(* IEC 61131-3 sources: laba_2_/Libraries/Acp10_MC (part 3) *)

FUNCTION_BLOCK MC_BR_OffsetVelocity (*adds a velocity offset to the velocity of the slave axis*)
	VAR_INPUT
		Slave : UDINT; (*axis reference of the slave axis*)
		Enable : BOOL; (*enable the function block*)
		CyclicVelocity : REAL; (*additive velocity*)
		Acceleration : REAL; (*acceleration for reaching the additive velocity*)
		AdvancedParameters : MC_ADV_OFFSETVELOCITY_REF; (*structure for using additional functions*)
	END_VAR
	VAR_OUTPUT
		Active : BOOL; (*a velocity offset can be executed*)
		Busy : BOOL; (*function block is not finished*)
		Error : BOOL; (*error occurred in FB*)
		ErrorID : UINT; (*error number*)
		VelocityAttained : BOOL; (*additive velocity offset reached*)
		ActualShiftValue : REAL; (*current value of velocity offset on the drive*)
	END_VAR
	VAR
		C_Slave : UDINT; (*internal variable*)
		IS : MC_0127_IS_TYP; (*internal variable*)
	END_VAR
END_FUNCTION_BLOCK

FUNCTION_BLOCK MC_BR_OffsetZone (*adds an offset to the position of the slave axis*)
	VAR_INPUT
		Slave : UDINT; (*axis reference of the slave axis*)
		Enable : BOOL; (*enable the function block*)
		InitData : BOOL; (*initialize the input data*)
		Shift : REAL; (*offset shift value*)
		Velocity : REAL; (*velocity for reaching the offset shift*)
		Acceleration : REAL; (*acceleration for reaching the offset shift*)
		ZoneStartPosition : REAL; (*start position of the offset shift zone*)
		ZoneEndPosition : REAL; (*end position of the offset shift zone*)
		AdvancedParameters : MC_ADV_OFFSETZONE_REF; (*structure for using additional functions*)
	END_VAR
	VAR_OUTPUT
		Active : BOOL; (*a offset shift can be executed*)
		Busy : BOOL; (*function block is not finished*)
		Error : BOOL; (*error occurred in FB*)
		ErrorID : UINT; (*error number*)
		ShiftAttained : BOOL; (*offset shift executed*)
		DataInitialized : BOOL; (*input data initialized*)
		ActualShiftValue : REAL; (*current value of shift on the drive*)
	END_VAR
	VAR
		C_Slave : UDINT; (*internal variable*)
		IS : MC_0128_IS_TYP; (*internal variable*)
	END_VAR
END_FUNCTION_BLOCK

FUNCTION_BLOCK MC_BR_GetParIDInfo (*determines data type and data length of a ParID*)
	VAR_INPUT
		Execute : BOOL; (*determine ParID information at rising edge*)
		ParID : UINT; (*ParID of which the information should be determined*)
	END_VAR
	VAR_OUTPUT
		Done : BOOL; (*command executed*)
		Busy : BOOL; (*function block is not finished*)
		Error : BOOL; (*error occurred in FB*)
		ErrorID : UINT; (*error number*)
		ParIDInfo : MC_PARID_INFO_REF; (*information about ParID*)
	END_VAR
	VAR
		IS : MC_0106_IS_TYP; (*intern variable*)
	END_VAR
END_FUNCTION_BLOCK

FUNCTION_BLOCK MC_BR_ParTrace (*controls the parameter trace*)
	VAR_INPUT
		Execute : BOOL; (*execute command at rising edge*)
		Command : UINT; (*select the command for the trace*)
		Configuration : MC_PARTRACECONFIG_REF; (*FB configuration*)
	END_VAR
	VAR_OUTPUT
		Done : BOOL; (*command executed*)
		Busy : BOOL; (*function block is not finished*)
		Error : BOOL; (*error occurred in FB*)
		ErrorID : UINT; (*error number*)
		ErrorRecord : MC_ERRORRECORD_REF; (*error messages that can occur after executing the command*)
	END_VAR
	VAR
		IS : MC_0080_IS_TYP; (*intern variable*)
	END_VAR
END_FUNCTION_BLOCK

FUNCTION_BLOCK MC_BR_ParTraceConfig (*load and save axis trace configuration*)
	VAR_INPUT
		Execute : BOOL; (*execute command at rising edge*)
		Command : UINT; (*select the command for the trace*)
		AdrTraceConfig : UDINT; (*adress of axis trace configuration*)
		DataObject : MC_DATOBJ_REF; (*data object parameters*)
	END_VAR
	VAR_OUTPUT
		Done : BOOL; (*command executed*)
		Busy : BOOL; (*function block is not finished*)
		Error : BOOL; (*error occurred in FB*)
		ErrorID : UINT; (*error number*)
		ErrorRecord : MC_ERRORRECORD_REF; (*error messages that can occur after executing the command*)
	END_VAR
	VAR
		IS : MC_0102_IS_TYP; (*intern variable*)
	END_VAR
END_FUNCTION_BLOCK

FUNCTION_BLOCK MC_BR_Phasing (*causes a phase shift in the master position of the slave axis*)
	VAR_INPUT
		Slave : UDINT; (*axis reference of the slave axis*)
		Enable : BOOL; (*enable the function block*)
		InitData : BOOL; (*initialize the input data*)
		PerformVelocityControl : BOOL; (*enable the phase shift*)
		Shift : REAL; (*phase shift value*)
		Velocity : REAL; (*velocity for reaching the phase shift*)
		Acceleration : REAL; (*acceleration for reaching the phase shift*)
		ApplicationDistance : REAL; (*distance within which the phase shift occurs*)
		ApplicationMode : UINT; (*basis for movement profile*)
		ShiftMode : UINT; (*definition of how the value on the "Shift" input should be used*)
		AdvancedParameters : MC_ADVANCEDSHIFTPAR_REF; (*structure for using additional functions*)
	END_VAR
	VAR_OUTPUT
		Active : BOOL; (*a phase shift can be executed*)
		Busy : BOOL; (*function block is not finished*)
		Error : BOOL; (*error occurred in FB*)
		ErrorID : UINT; (*error number*)
		ShiftAttained : BOOL; (*phase shift executed*)
		DataInitialized : BOOL; (*input data initialized*)
		ActualShiftValue : REAL; (*current value of shift on the drive*)
	END_VAR
	VAR
		C_Slave : UDINT; (*internal variable*)
		C_InitData : BOOL; (*internal variable*)
		C_PerformVelocityControl : BOOL; (*internal variable*)
		C_Shift : DINT; (*internal variable*)
		C_Velocity : REAL; (*internal variable*)
		C_Acceleration : REAL; (*internal variable*)
		C_ApplicationDistance : DINT; (*internal variable*)
		C_ApplicationMode : UINT; (*internal variable*)
		C_SelectedMaster : UINT; (*internal variable*)
		C_ShiftMode : UINT; (*internal variable*)
		C_AdvancedParameters : MC_ADVANCEDSHIFTPAR_REF; (*internal variable*)
		C_Active : BOOL; (*internal variable*)
		C_Busy : BOOL; (*internal variable*)
		C_Error : BOOL; (*internal variable*)
		C_ErrorID : UINT; (*internal variable*)
		CC_ErrorID : UINT; (*internal variable*)
		C_ShiftAttained : BOOL; (*internal variable*)
		C_DataInitialized : BOOL; (*internal variable*)
		C_AxisState : UINT; (*internal variable*)
		NextState : USINT; (*internal variable*)
		state : USINT; (*internal variable*)
		LockID : USINT; (*internal variable*)
		LockIDPar : USINT; (*internal variable*)
		Factor : UDINT; (*internal variable*)
		RtN : REAL; (*internal variable*)
		VarIndex : UINT; (*internal variable*)
		MpgenIndex : UINT; (*internal variable*)
		C_MpgenStatus : USINT; (*internal variable*)
		MpgenStatusOffset : UINT; (*internal variable*)
		MpgenStatusRecIndex : USINT; (*internal variable*)
		Reserve : USINT; (*internal variable*)
		MpgenValueOffset : UINT; (*internal variable*)
		MpgenValueRecIndex : USINT; (*internal variable*)
		FbID : USINT; (*internal variable*)
		InitDataActive : BOOL; (*internal variable*)
	END_VAR
END_FUNCTION_BLOCK

FUNCTION_BLOCK MC_BR_MechPosDeviationComp (*handles mechanics position deviation compensation*)
	VAR_INPUT
		Axis : UDINT; (*axis reference*)
		Enable : BOOL; (*as long as Enable is TRUE the FB is active*)
		Parameters : MC_MPDC_PARAM_REF; (*parameters for mechanics position deviation compensation*)
		AdvancedParameters : MC_ADV_MPDC_REF; (*advanced parameters for mechanics deviation position compensation*)
	END_VAR
	VAR_OUTPUT
		Active : BOOL; (*if set, the mechanics deviation position compensation is active*)
		Busy : BOOL; (*function block is not finished*)
		Error : BOOL; (*error occurred in FB*)
		ErrorID : UINT; (*error number*)
		AdvancedInfo : MC_ADV_INFO_MPDC_REF; (*structure with additional information*)
	END_VAR
	VAR
		C_Axis : UDINT; (*internal variable*)
		IS : MC_0147_IS_TYP; (*internal structure*)
	END_VAR
END_FUNCTION_BLOCK

FUNCTION_BLOCK MC_BR_PowerMeter (*executes the evaluation of the powerdata of a PSM*)
	VAR_INPUT
		Axis : UDINT; (*axis reference*)
		Enable : BOOL; (*as long as Enable is TRUE the power evaluation is active*)
		Mode : USINT; (*choose the mode for the power evaluation*)
		IntervalTime : UINT; (*duration of the interval*)
		RestartInterval : BOOL; (*a new interval is startet at rising edge of this input*)
		EventInput : MC_BR_EVINPUT_REF; (*if this is used, the Trigger input will not be considered*)
	END_VAR
	VAR_OUTPUT
		Valid : BOOL; (*if set, the data on Output PowerData are valid*)
		Busy : BOOL; (*function block is not finished*)
		Error : BOOL; (*error occurred in FB*)
		ErrorID : UINT; (*error number*)
		PowerData : MC_POWERDATA_REF; (*structure for the power data*)
		MissedIntervals : UINT; (*count of missed intervalls*)
	END_VAR
	VAR
		C_Axis : UDINT; (*internal variable*)
		IS : MC_0089_IS_TYP; (*internal structure*)
	END_VAR
END_FUNCTION_BLOCK

FUNCTION_BLOCK MC_BR_ReadAutPosition (*reads the cam profile automat position*)
	VAR_INPUT
		Axis : UDINT; (*axis reference*)
		Execute : BOOL; (*automat position is read at rising edge*)
	END_VAR
	VAR_OUTPUT
		Done : BOOL; (*reading automat position is finished*)
		Busy : BOOL; (*function block is not finished*)
		Error : BOOL; (*error occurred in FB*)
		ErrorID : UINT; (*error number*)
		AutPosition : REAL; (*automat position*)
	END_VAR
	VAR
		C_Axis : UDINT; (*internal variable*)
		C_Execute : BOOL; (*internal variable*)
		C_Done : BOOL; (*internal variable*)
		C_Error : BOOL; (*internal variable*)
		C_ErrorID : UINT; (*internal variable*)
		LockIDPar : USINT; (*internal variable*)
		Reserve1 : USINT; (*internal variable*)
		C_AutPosition : DINT; (*internal variable*)
		C_DataAddress : UDINT; (*internal variable*)
		state : USINT; (*internal variable*)
	END_VAR
END_FUNCTION_BLOCK

FUNCTION_BLOCK MC_BR_ReadAxisError (*reads and acknowledges an axis error record and reads the error text*)
	VAR_INPUT
		Axis : UDINT; (*axis reference*)
		Enable : BOOL; (*read error record/text*)
		Acknowledge : BOOL; (*acknowledge current axis error*)
		Mode : UINT; (*operating mode of FB*)
		Configuration : MC_ERRORTEXTCONFIG_REF; (*FB configuration*)
	END_VAR
	VAR_OUTPUT
		Valid : BOOL; (*if set, the data of the other outputs is valid*)
		Busy : BOOL; (*function block is not finished*)
		Error : BOOL; (*error occurred in FB*)
		ErrorID : UINT; (*error number*)
		ErrorRecordAvailable : BOOL; (*a new error record is available*)
		ErrorRecord : MC_ERRORRECORD_REF; (*detailed axis error information*)
		FunctionBlockErrorCount : UINT; (*number of not acknowledged function block errors*)
		AxisErrorCount : UINT; (*number of not acknowledged axis errors*)
		AxisWarningCount : UINT; (*number of not acknowledged axis warnings*)
	END_VAR
	VAR
		C_Axis : UDINT; (*internal variable*)
		IS : MC_0105_IS_TYP; (*internal variable*)
	END_VAR
END_FUNCTION_BLOCK

FUNCTION_BLOCK MC_BR_ReadCyclicPosition (*read the position of an axis cyclically*)
	VAR_INPUT
		Axis : UDINT; (*axis reference*)
		Enable : BOOL; (*as long as Enable is TRUE the cyclic position is read from the axis*)
		ParID : UINT; (*ParID that is read cyclically, 0... set position*)
	END_VAR
	VAR_OUTPUT
		Valid : BOOL; (*position is beeing read from the axis*)
		Busy : BOOL; (*function block is not finished*)
		Error : BOOL; (*error occurred in FB*)
		ErrorID : UINT; (*error number*)
		CyclicPosition : MC_CYCLIC_POSITION; (*cyclic position that is read from the axis*)
	END_VAR
	VAR
		C_Axis : UDINT; (*internal variable*)
		IS : MC_0082_IS_TYP; (*internal variable*)
	END_VAR
END_FUNCTION_BLOCK

FUNCTION_BLOCK MC_BR_ReadDriveStatus (*checks the status of a drive*)
	VAR_INPUT
		Axis : UDINT; (*axis reference*)
		Enable : BOOL; (*when set the status is read*)
		AdrDriveStatus : UDINT; (*address of the structur where the status is written on*)
	END_VAR
	VAR_OUTPUT
		Valid : BOOL; (*output of FB is valid*)
		Busy : BOOL; (*function block is not finished*)
		Error : BOOL; (*error occurred in FB*)
		ErrorID : UINT; (*error number*)
	END_VAR
	VAR
		C_Axis : UDINT; (*internal variable*)
		state : USINT; (*internal variable*)
		C_Error : BOOL; (*internal variable*)
		C_ErrorID : UINT; (*internal variable*)
		C_AdrDriveStatus : UDINT; (*internal variable*)
	END_VAR
END_FUNCTION_BLOCK

FUNCTION_BLOCK MC_BR_ReadNetTraceStatus (*determines the current status of the network command trace*)
	VAR_INPUT
		Enable : BOOL; (*the status of the network command trace is read as long as the input is enabled*)
		Configuration : MC_NETTRACECONFIG_REF; (*FB configuration. Only the element "NetTrace" is evaluated*)
	END_VAR
	VAR_OUTPUT
		Valid : BOOL; (*the status information is valid*)
		Busy : BOOL; (*function block is not finished*)
		Error : BOOL; (*error occurred in FB*)
		ErrorID : UINT; (*error number*)
		TraceState : UINT; (*status of the NWCT*)
	END_VAR
	VAR
		C_ErrorID : UINT; (*internal variable*)
		C_Error : BOOL; (*internal variable*)
		state : USINT; (*internal variable*)
	END_VAR
END_FUNCTION_BLOCK

FUNCTION_BLOCK MC_BR_ReadParID (*reads a ParID from the specified axis*)
	VAR_INPUT
		Axis : UDINT; (*axis reference*)
		Execute : BOOL; (*read data at rising edge*)
		ParID : UINT; (*number of the parameter ID to read*)
		DataAddress : UDINT; (*address of the user variable*)
		DataType : UINT; (*data type of the user variable*)
	END_VAR
	VAR_OUTPUT
		Done : BOOL; (*value of ParID has been copied to the user variable*)
		Busy : BOOL; (*function block is not finished*)
		Error : BOOL; (*error occurred in function block*)
		ErrorID : UINT; (*error number*)
	END_VAR
	VAR
		C_Axis : UDINT; (*internal variable*)
		C_Execute : BOOL; (*internal variable*)
		C_ParID : UINT; (*internal variable*)
		LockIDPar : USINT; (*internal variable*)
		Reserve1 : USINT; (*internal variable*)
		C_DataAddress : UDINT; (*internal variable*)
		Reserve2 : UDINT; (*internal variable*)
		C_DataType : UINT; (*internal variable*)
		C_Done : BOOL; (*internal variable*)
		C_Error : BOOL; (*internal variable*)
		C_ErrorID : UINT; (*internal variable*)
		state : USINT; (*internal variable*)
	END_VAR
END_FUNCTION_BLOCK

FUNCTION_BLOCK MC_BR_ReadParIDText (*reads a ParID from the specified axis in text format*)
	VAR_INPUT
		Axis : UDINT; (*axis reference*)
		Execute : BOOL; (*read data at rising edge*)
		ParID : UINT; (*number of the parameter ID to read*)
	END_VAR
	VAR_OUTPUT
		Done : BOOL; (*value of ParID has been read*)
		Busy : BOOL; (*function block is not finished*)
		Error : BOOL; (*error occurred in function block*)
		ErrorID : UINT; (*error number*)
		DataText : STRING[33]; (*value of ParID in text format *)
	END_VAR
	VAR
		C_Axis : UDINT; (*internal variable*)
		C_Execute : BOOL; (*internal variable*)
		C_ParID : UINT; (*internal variable*)
		LockIDPar : USINT; (*internal variable*)
		C_Done : BOOL; (*internal variable*)
		C_Error : BOOL; (*internal variable*)
		C_ErrorID : UINT; (*internal variable*)
		state : USINT; (*internal variable*)
	END_VAR
END_FUNCTION_BLOCK

FUNCTION_BLOCK MC_BR_ReadParList (*read a parameter list*)
	VAR_INPUT
		Axis : UDINT; (*axis reference*)
		Execute : BOOL; (*read parameter list at rising edge*)
		DataAddress : UDINT; (*address of the parameter list*)
	END_VAR
	VAR_OUTPUT
		Done : BOOL; (*transfer completed*)
		Busy : BOOL; (*function block is not finished*)
		Error : BOOL; (*error occurred in FB*)
		ErrorID : UINT; (*error number*)
	END_VAR
	VAR
		LockIDPar : USINT; (*internal variable*)
		C_Error : BOOL; (*internal variable*)
		C_ErrorID : UINT; (*internal variable*)
		C_Axis : UDINT; (*internal variable*)
		C_DataAddress : UDINT; (*internal variable*)
		C_Done : BOOL; (*internal variable*)
		state : USINT; (*internal variable*)
	END_VAR
END_FUNCTION_BLOCK

FUNCTION_BLOCK MC_BR_ReadParTraceStatus (*determines the current status of the axis trace*)
	VAR_INPUT
		Enable : BOOL; (*the status of the axis trace is read as long as the input is enabled*)
		Configuration : MC_PARTRACECONFIG_REF; (*FB configuration. Only the element "ParTrace" is evaluated*)
	END_VAR
	VAR_OUTPUT
		Valid : BOOL; (*the status information is valid*)
		Busy : BOOL; (*function block is not finished*)
		Error : BOOL; (*error occurred in FB*)
		ErrorID : UINT; (*error number*)
		TraceState : UINT; (*status of the trace*)
	END_VAR
	VAR
		C_ErrorID : UINT; (*internal variable*)
		C_Error : BOOL; (*internal variable*)
		state : USINT; (*internal variable*)
	END_VAR
END_FUNCTION_BLOCK

FUNCTION_BLOCK MC_BR_ReceiveParIDOnPLC (*initializes receiving of a ParID on the PLC*)
	VAR_INPUT
		Axis : UDINT; (*axis reference*)
		Enable : BOOL; (*as long as Enable is TRUE the ParID is read from the axis*)
		ParID : UINT; (*ParID that is read cyclically*)
		SendChannel : USINT; (*send channel on which the ParID is sent*)
		Mode : USINT; (*convertion of ParID-value into PLCopen-units can be activated*)
	END_VAR
	VAR_OUTPUT
		Valid : BOOL; (*ParID is beeing read from the axis*)
		Busy : BOOL; (*function block is not finished*)
		Error : BOOL; (*error occurred in FB*)
		ErrorID : UINT; (*error number*)
		CyclicValue : MC_CYCLIC_VALUE_REF; (*cyclic ParID value that is read from the axis*)
	END_VAR
	VAR
		C_Axis : UDINT; (*internal variable*)
		IS : MC_0113_IS_TYP; (*internal variable*)
	END_VAR
END_FUNCTION_BLOCK

FUNCTION_BLOCK MC_BR_ResetAutPar (*initializes the general parameters of the cam automat*)
	VAR_INPUT
		Axis : UDINT; (*axis reference*)
		Execute : BOOL; (*set parameter to default values at rising edge*)
		GlobalParams : USINT; (*selection of the global parameter*)
		StateIndex : USINT; (*selection of the automat state*)
	END_VAR
	VAR_OUTPUT
		Done : BOOL; (*automat parameters set to default values*)
		Busy : BOOL; (*function block not finished*)
		Error : BOOL; (*error occurred in FB*)
		ErrorID : UINT; (*error number*)
	END_VAR
	VAR
		C_Axis : UDINT; (*internal variable*)
		IS : MC_0136_IS_TYP; (*internal variable*)
	END_VAR
END_FUNCTION_BLOCK

FUNCTION_BLOCK MC_BR_SaveAxisPar (*writes the axis parameters in the axis data structure*)
	VAR_INPUT
		Axis : UDINT; (*axis reference*)
		Execute : BOOL; (*write axis parameter from the axis structure to a init parameter module at rising edge*)
		DataObjectName : STRING[12]; (*name of the init parameter module*)
	END_VAR
	VAR_OUTPUT
		Done : BOOL; (*saving the data is finished*)
		Busy : BOOL; (*function block is not finished*)
		Error : BOOL; (*error occurred in FB*)
		ErrorID : UINT; (*error number*)
		DataObjectIdent : UDINT; (*init parameter module data object ID for the function blocks in the DataObj library*)
	END_VAR
	VAR
		C_Axis : UDINT;
		C_DataObjectName : STRING[12]; (*internal variable*)
		state : USINT; (*internal variable*)
		LockIDPar : USINT; (*internal variable*)
		C_ErrorID : UINT; (*internal variable*)
		C_Error : BOOL; (*internal variable*)
		pInit : REFERENCE TO USINT; (*internal variable*)
		pError : REFERENCE TO USINT; (*internal variable*)
	END_VAR
END_FUNCTION_BLOCK

FUNCTION_BLOCK MC_BR_SaveCamProfileObj (*saves the data of a cam profile into a data module*)
	VAR_INPUT
		Execute : BOOL; (*save the cam profile at rising edge*)
		DataObjectName : STRING[12]; (*name for the data module in which the cam profile is saved*)
		DataAddress : UDINT; (*address of the cam profile data*)
		DataObjectVersion : UINT; (*version for the data module*)
	END_VAR
	VAR_OUTPUT
		Done : BOOL; (*data module was saved*)
		Busy : BOOL; (*function block is not finished*)
		Error : BOOL; (*error occurred in FB*)
		ErrorID : UINT; (*error number*)
		ErrorRecord : MC_ERRORRECORD_REF; (*error messages that can occur after executing the command*)
		DataObjectIdent : UDINT; (*ident of the data module*)
	END_VAR
	VAR
		IS : MC_0116_IS_TYP; (*internal variable*)
	END_VAR
END_FUNCTION_BLOCK

FUNCTION_BLOCK MC_BR_SetHardwareInputs (*forces the hardware inputs*)
	VAR_INPUT
		Axis : UDINT; (*axis reference*)
		Enable : BOOL; (*set the status of the hardware inputs as long as the input is enabled*)
		HomeSwitch : BOOL; (*if TRUE the reference hardware input is activated*)
		PosHWSwitch : BOOL; (*if TRUE the positive limit switch input is activated*)
		NegHWSwitch : BOOL; (*if TRUE the negative limit switch input is activated*)
		Trigger1 : BOOL; (*if TRUE the trigger1 input is activated*)
		Trigger2 : BOOL; (*if TRUE the trigger2 input is activated*)
	END_VAR
	VAR_OUTPUT
		Active : BOOL; (*function block is active and waits for changes on the inputs*)
		Busy : BOOL; (*function block is not finished*)
		Error : BOOL; (*error occurred in FB*)
		ErrorID : UINT; (*error number*)
		InputsSet : BOOL; (*the actual input status was transferred*)
	END_VAR
	VAR
		C_Axis : UDINT; (*internal variable*)
		IS : MC_0108_IS_TYP; (*internal variable*)
	END_VAR
END_FUNCTION_BLOCK

FUNCTION_BLOCK MC_BR_SetupController (*starts a controller setup and saves the parameters*)
	VAR_INPUT
		Axis : UDINT; (*axis reference*)
		Execute : BOOL; (*starts the command action at rising edge*)
		Command : UINT; (*choose the command for the setup*)
		Configuration : MC_SETUP_CONTROLLER_CFG_REF; (*FB-Configuration*)
	END_VAR
	VAR_OUTPUT
		Done : BOOL; (*command successfully completed*)
		Busy : BOOL; (*function block is not finished*)
		CommandAborted : BOOL; (*function block is aborted by another command*)
		Error : BOOL; (*error occurred in FB*)
		ErrorID : UINT; (*error number*)
		SetupOutput : MC_SETUP_OUTPUT_REF; (*structure for output values*)
	END_VAR
	VAR
		C_Axis : UDINT; (*internal variable*)
		IS : MC_0090_IS_TYP; (*internal variable*)
	END_VAR
END_FUNCTION_BLOCK

FUNCTION_BLOCK MC_BR_SetupFromParTabObj (*starts a setup with parameter from an ACOPOS parameter table*)
	VAR_INPUT
		Axis : UDINT; (*axis reference*)
		Execute : BOOL; (*starts the commanded action at rising edge*)
		Command : UINT; (*choose the command for the setup*)
		DataObjectName : STRING[12]; (*name of the ACOPOS parameter table*)
	END_VAR
	VAR_OUTPUT
		Done : BOOL; (*command succesfully completed*)
		Busy : BOOL; (*function block is not finished*)
		CommandAborted : BOOL; (*function block is aborted by another command*)
		Error : BOOL; (*error occurred in FB*)
		ErrorID : UINT; (*error number*)
		SetupOutput : MC_SETUP_OUTPUT_REF; (*structure for output values*)
	END_VAR
	VAR
		C_Axis : UDINT; (*internal variable*)
		IS : MC_0145_IS_TYP; (*internal variable*)
	END_VAR
END_FUNCTION_BLOCK

FUNCTION_BLOCK MC_BR_SetupInductionMotor (*starts the motorsetup for an induction motor and saves the parameters*)
	VAR_INPUT
		Axis : UDINT; (*axis reference*)
		Execute : BOOL; (*starts the commanded action at rising edge*)
		Command : UINT; (*choose the command for the setup*)
		Configuration : MC_SETUP_IND_MOTOR_CFG_REF; (*FB-Configuration*)
	END_VAR
	VAR_OUTPUT
		Done : BOOL; (*command succesfully completed*)
		Busy : BOOL; (*function block is not finished*)
		CommandAborted : BOOL; (*function block is aborted by another command*)
		Error : BOOL; (*error occurred in FB*)
		ErrorID : UINT; (*error number*)
		SetupOutput : MC_SETUP_OUTPUT_REF; (*structure for output values*)
	END_VAR
	VAR
		C_Axis : UDINT; (*internal variable*)
		IS : MC_0088_IS_TYP; (*internal variable*)
	END_VAR
END_FUNCTION_BLOCK

FUNCTION_BLOCK MC_BR_SetupIsqRipple (*starts the setup for isq ripple compensation  and saves the parameters*)
	VAR_INPUT
		Axis : UDINT; (*axis reference*)
		Execute : BOOL; (*starts the commanded action at rising edge*)
		Command : UINT; (*choose the command for the setup*)
		Configuration : MC_SETUP_ISQ_RIPPLE_CFG_REF; (*FB-Configuration*)
	END_VAR
	VAR_OUTPUT
		Done : BOOL; (*command successfully completed*)
		Busy : BOOL; (*function block is not finished*)
		CommandAborted : BOOL; (*function block is aborted by another command*)
		Error : BOOL; (*error occurred in FB*)
		ErrorID : UINT; (*error number*)
		SetupOutput : MC_SETUP_OUTPUT_REF; (*structure for the output values*)
	END_VAR
	VAR
		C_Axis : UDINT; (*internal variable*)
		IS : MC_0101_IS_TYP; (*internal variable*)
	END_VAR
END_FUNCTION_BLOCK

FUNCTION_BLOCK MC_BR_SetupMotorPhasing (*starts a phasing setup and saves the parameters*)
	VAR_INPUT
		Axis : UDINT; (*axis reference*)
		Execute : BOOL; (*starts the commanded action at rising edge*)
		Command : UINT; (*choose the command for the setup*)
		Configuration : MC_SETUP_MOTOR_PHA_CFG_REF; (*FB-Configuration*)
	END_VAR
	VAR_OUTPUT
		Done : BOOL; (*command successfully completed*)
		Busy : BOOL; (*function block is not finished*)
		CommandAborted : BOOL; (*function block is aborted by another command*)
		Error : BOOL; (*error occurred in FB*)
		ErrorID : UINT; (*error number *)
		SetupOutput : MC_SETUP_OUTPUT_REF; (*structure for output values*)
		SetupResult : MC_SETUP_PHASING_RESULT_REF; (*structure for results of the setup*)
	END_VAR
	VAR
		C_Axis : UDINT; (*internal variable*)
		IS : MC_0097_IS_TYP; (*internal variable*)
	END_VAR
END_FUNCTION_BLOCK

FUNCTION_BLOCK MC_BR_SetupSynchronMotor (*starts the motorsetup for a synchron motor and saves the parameters*)
	VAR_INPUT
		Axis : UDINT; (*axis reference*)
		Execute : BOOL; (*starts the commanded action at rising edge*)
		Command : UINT; (*choose the command for the setup*)
		Configuration : MC_SETUP_SYNC_MOTOR_CFG_REF; (*FB-Configuration*)
	END_VAR
	VAR_OUTPUT
		Done : BOOL; (*command successfully completed*)
		Busy : BOOL; (*function block is not finished*)
		CommandAborted : BOOL; (*function block is aborted by another command*)
		Error : BOOL; (*error occurred in FB*)
		ErrorID : UINT; (*error number*)
		SetupOutput : MC_SETUP_OUTPUT_REF; (*structure for output values*)
	END_VAR
	VAR
		C_Axis : UDINT; (*internal variable*)
		IS : MC_0129_IS_TYP; (*internal variable*)
	END_VAR
END_FUNCTION_BLOCK

FUNCTION_BLOCK MC_BR_Simulation (*turns on or off simulation mode for a drive*)
	VAR_INPUT
		Axis : UDINT; (*axis reference*)
		Execute : BOOL; (*switch simulation mode on or off at rising edge*)
		SimulationCommand : UINT; (*choose if switch on or off simulation mode*)
	END_VAR
	VAR_OUTPUT
		Done : BOOL; (*simulation mode is on or off*)
		Busy : BOOL; (*function block is not finished*)
		Error : BOOL; (*error occurred in FB*)
		ErrorID : UINT; (*error number*)
	END_VAR
	VAR
		C_Axis : UDINT; (*internal variable*)
		IS : MC_0071_IS_TYP; (*internal variable*)
	END_VAR
END_FUNCTION_BLOCK

FUNCTION_BLOCK MC_BR_TouchProbe (*saves the values of ParIDs when a specified event occurs*)
	VAR_INPUT
		Axis : UDINT; (*axis reference*)
		TriggerInput : MC_BR_TRIGGER_REF; (*input that is used as event source*)
		Enable : BOOL; (*as long as enable is TRUE, a value is saved every time a trigger event occurs*)
		Period : REAL; (*interval between two expected trigger positions*)
		PeriodChange : REAL; (*if no valid event occurs within an interval, the window is shifted by the value of Period*)
		ExpectedValue : REAL; (*expected position of the trigger event within the Period*)
		WindowNegative : REAL; (*range before the expected position in which the trigger signal may occur*)
		WindowPositive : REAL; (*range after the expected position in which the trigger signal may occur*)
		Mode : UINT; (*the way the FB works can be determined with this input*)
	END_VAR
	VAR_OUTPUT
		Active : BOOL; (*waits for a trigger event*)
		Busy : BOOL; (*function block is not finished*)
		Error : BOOL; (*error occured in FB*)
		ErrorID : UINT; (*error number*)
		RecordedPeriodicValue : REAL; (*result value within the configured period*)
		RecordedValue : DINT; (*result value*)
		DeltaExpectedValue : REAL; (*deviation: expected position - result value*)
		ProbeCounter : UDINT; (*number of valid trigger events since "Enable" was set to TRUE*)
		MissedTriggers : UDINT; (*number of invalid or missing trigger events since "Enable" was set to TRUE*)
	END_VAR
	VAR
		C_Axis : UDINT; (*internal variable*)
		C_TriggerInput : MC_BR_TRIGGER_REF; (*internal variable*)
		C_Period : DINT; (*internal variable*)
		C_PeriodChange : DINT; (*internal variable*)
		C_ExpectedValue : DINT; (*internal variable*)
		C_WindowNegative : DINT; (*internal variable*)
		C_WindowPositive : DINT; (*internal variable*)
		C_Mode : UINT; (*internal variable*)
		C_Active : BOOL; (*internal variable*)
		C_Busy : BOOL; (*internal variable*)
		C_Error : BOOL; (*internal variable*)
		C_ErrorID : UINT; (*internal variable*)
		C_RecordedPeriodicValue : REAL; (*internal variable*)
		C_RecordedValue : DINT; (*internal variable*)
		C_DeltaExpectedValue : REAL; (*internal variable*)
		C_ProbeCounter : UDINT; (*internal variable*)
		C_MissedTriggers : UDINT; (*internal variable*)
		PeriodOffset : DINT; (*internal variable*)
		LatchValue : DINT; (*internal variable*)
		LatchDeltaIv : DINT; (*internal variable*)
		NewValue : BOOL; (*internal variable*)
		state : USINT; (*internal variable*)
		NextState : USINT; (*internal variable*)
		DataTyp : UINT; (*internal variable*)
		LockIDPar : USINT; (*internal variable*)
		LockID : USINT; (*internal variable*)
		ActualPosition : DINT; (*internal variable*)
		LatchIndex : UINT; (*internal variable*)
		BitIndex : UINT; (*internal variable*)
		BitValueOffset : UINT; (*internal variable*)
		BitValueRecIndex : USINT; (*internal variable*)
		SptID : USINT; (*internal variable*)
		UpdatePeriod : BOOL; (*internal variable*)
		UseAxisPeriod : BOOL; (*internal variable*)
	END_VAR
END_FUNCTION_BLOCK

FUNCTION_BLOCK MC_BR_VelocityControl (*sends cyclic speed set value for velocity control*)
	VAR_INPUT
		Axis : UDINT; (*axis reference*)
		Enable : BOOL; (*when set the FB will activate torque control*)
		CyclicVelocity : REAL; (*Parameter input for set speed*)
		CyclicVelocityCorrection : REAL; (*Parameter input for additive set speed*)
		CyclicTorque : REAL; (*Parameter input for limit or additive torque*)
		TorqueMode : USINT; (*Mode setting (limit or additive torque)*)
		Acceleration : REAL; (*Value of maximum acceleration*)
		Deceleration : REAL; (*Value of maximum deceleration*)
		SctrlKv : REAL; (*Value of proportional part of speed controller*)
		SctrlTn : REAL; (*Value of integral part of speed controller*)
		InitSctrl : BOOL; (*Command for downloading values for sctrl*)
	END_VAR
	VAR_OUTPUT
		Active : BOOL; (*Functionality of FB enabled*)
		Busy : BOOL; (*Function Block is not finished*)
		CommandAborted : BOOL; (*FB was aborted from MC_Power or an Error*)
		Error : BOOL; (*Error occured in FB*)
		ErrorID : UINT; (*PLCopen error number*)
		SctrlInitialized : BOOL; (*Parameters to speed controller downloaded*)
	END_VAR
	VAR
		C_Axis : UDINT; (*internal variable*)
		IS : MC_0095_IS_TYP; (*internal structure*)
	END_VAR
END_FUNCTION_BLOCK

FUNCTION_BLOCK MC_BR_WriteParID (*writes a ParID to specified axis*)
	VAR_INPUT
		Axis : UDINT; (*axis reference*)
		Execute : BOOL; (*write data at rising edge*)
		ParID : UINT; (*number of the parameter ID to write*)
		DataAddress : UDINT; (*address of the user variable*)
		DataType : UINT; (*data type of user variable*)
	END_VAR
	VAR_OUTPUT
		Done : BOOL; (*value of the user variable has been copied to the ParID*)
		Busy : BOOL; (*parameter write is in progress*)
		Error : BOOL; (*error occurred in FB*)
		ErrorID : UINT; (*error number*)
	END_VAR
	VAR
		C_Axis : UDINT; (*internal variable*)
		C_Execute : BOOL; (*internal variable*)
		C_ParID : UINT; (*internal variable*)
		LockIDPar : USINT; (*internal variable*)
		Reserve1 : USINT; (*internal variable*)
		C_DataAddress : UDINT; (*internal variable*)
		Reserve2 : UDINT; (*internal variable*)
		C_DataType : UINT; (*internal variable*)
		C_Done : BOOL; (*internal variable*)
		C_Error : BOOL; (*internal variable*)
		C_ErrorID : UINT; (*internal variable*)
		state : USINT; (*internal variable*)
	END_VAR
END_FUNCTION_BLOCK

FUNCTION_BLOCK MC_BR_WriteParIDText (*writes a ParID from the specified axis in text format*)
	VAR_INPUT
		Axis : UDINT; (*axis reference*)
		Execute : BOOL; (*write data at rising edge*)
		ParID : UINT; (*number of the parameter ID to write*)
		DataText : STRING[33]; (*value of ParID in text format *)
	END_VAR
	VAR_OUTPUT
		Done : BOOL; (*value of ParID has been written*)
		Busy : BOOL; (*function block is not finished*)
		Error : BOOL; (*error occurred in function block*)
		ErrorID : UINT; (*error number*)
	END_VAR
	VAR
		C_Axis : UDINT; (*internal variable*)
		C_Execute : BOOL; (*internal variable*)
		C_ParID : UINT; (*internal variable*)
		LockIDPar : USINT; (*internal variable*)
		C_Done : BOOL; (*internal variable*)
		C_Error : BOOL; (*internal variable*)
		C_ErrorID : UINT; (*internal variable*)
		state : USINT; (*internal variable*)
	END_VAR
END_FUNCTION_BLOCK

FUNCTION_BLOCK MC_CamIn (*engages a cam coupling between master and slave axis*)
	VAR_INPUT
		Master : UDINT; (*axis reference of the master axis*)
		Slave : UDINT; (*axis reference of the slave axis*)
		Execute : BOOL; (*start at rising edge*)
		MasterOffset : REAL; (*offset on master axis*)
		SlaveOffset : REAL; (*offset on slave axis*)
		MasterScaling : REAL; (*factor for the master profile*)
		SlaveScaling : REAL; (*factor for the slave profile*)
		StartMode : USINT; (*start mode*)
		CamTableID : USINT; (*identifier of cam table*)
		MasterParID : UINT; (*use this ParID instead of the set position*)
	END_VAR
	VAR_OUTPUT
		InSync : BOOL; (*cam is engaged for the first time*)
		Busy : BOOL; (*function block is not finished*)
		CommandAborted : BOOL; (*function block aborted by another command*)
		Error : BOOL; (*error occurred in FB*)
		ErrorID : UINT; (*error number*)
		EndOfProfile : BOOL; (*pulsed output signaling the cyclic end of the cam profile*)
	END_VAR
	VAR
		LockID : USINT; (*internal variable*)
		LockIDPar : USINT; (*internal variable*)
		LockIDInSync : USINT; (*internal variable*)
		C_Execute : BOOL; (*internal variable*)
		C_Master : UDINT; (*internal variable*)
		C_Slave : UDINT; (*internal variable*)
		C_MasterOffset : DINT; (*internal variable*)
		C_SlaveOffset : DINT; (*internal variable*)
		C_MasterScaling : DINT; (*internal variable*)
		C_SlaveScaling : DINT; (*internal variable*)
		C_CamTableID : UINT; (*internal variable*)
		C_StartMode : USINT; (*internal variable*)
		C_Periodic : BOOL; (*internal variable*)
		C_MasterParID : UINT; (*internal variable*)
		C_InSync : BOOL; (*internal variable*)
		C_CommandAborted : BOOL; (*internal variable*)
		C_ErrorID : UINT; (*internal variable*)
		C_Error : BOOL; (*internal variable*)
		C_EndOfProfile : BOOL; (*internal variable*)
		OldMaCamOffset : DINT; (*internal variable*)
		MaPosition : DINT; (*internal variable*)
		DataTyp : UINT; (*internal variable*)
		MpgenIndex : UINT; (*internal variable*)
		AutActualStateIndexOffset : UINT; (*internal variable*)
		AutActualStateIndexRecIndex : USINT; (*internal variable*)
		LockIDReceive : USINT; (*internal variable*)
		AutActualCamIndexOffset : UINT; (*internal variable*)
		AutActualCamIndexRecIndex : USINT; (*internal variable*)
		LockIDSend : USINT; (*internal variable*)
		AutMaCamOffsetOffset : UINT; (*internal variable*)
		AutMaCamOffsetRecIndex : USINT; (*internal variable*)
		LockIDMa : USINT; (*internal variable*)
		sendSlot : USINT; (*internal variable*)
		readSlot : USINT; (*internal variable*)
		state : USINT; (*internal variable*)
		MoveID : USINT; (*internal variable*)
		CC_ErrorID : UINT; (*internal variable*)
		oldMoveID : USINT; (*internal variable*)
	END_VAR
END_FUNCTION_BLOCK

FUNCTION_BLOCK MC_CamOut (*disengages the cam slave from the master axis*)
	VAR_INPUT
		Slave : UDINT; (*axis reference of the slave axis*)
		Execute : BOOL; (*start to disengage the slave from the master*)
	END_VAR
	VAR_OUTPUT
		Done : BOOL; (*disengaging complete*)
		Busy : BOOL; (*function block is not finished*)
		Error : BOOL; (*error occurred in FB*)
		ErrorID : UINT; (*error number*)
	END_VAR
	VAR
		C_Slave : UDINT; (*internal variable*)
		C_Execute : BOOL; (*internal variable*)
		C_Done : BOOL; (*internal variable*)
		C_Error : BOOL; (*internal variable*)
		C_ErrorID : UINT; (*internal variable*)
		state : USINT; (*internal variable*)
		LockIDPar : USINT; (*internal variable*)
		MoveID : USINT; (*internal variable*)
	END_VAR
END_FUNCTION_BLOCK

FUNCTION_BLOCK MC_CamTableSelect (*prepares the cam tables that will be used by the function block "MC_CamIn"*)
	VAR_INPUT
		Master : UDINT; (*axis reference of the master axis*)
		Slave : UDINT; (*axis reference of the slave axis*)
		CamTable : STRING[12]; (*name of the cam table*)
		Execute : BOOL; (*selection at rising edge*)
		Periodic : BOOL; (*select if periodic cam or non periodic cam*)
	END_VAR
	VAR_OUTPUT
		Done : BOOL; (*pre-selection done*)
		Busy : BOOL; (*function block is not finished*)
		Error : BOOL; (*error occurred in FB*)
		ErrorID : UINT; (*error number*)
		CamTableID : USINT; (*identifier of the cam table*)
	END_VAR
	VAR
		C_Master : UDINT; (*internal variable*)
		C_Slave : UDINT; (*internal variable*)
		C_CamTable : STRING[12]; (*internal variable*)
		Reserve : USINT; (*internal variable*)
		C_Periodic : BOOL; (*internal variable*)
		C_Error : BOOL; (*internal variable*)
		C_ErrorID : UINT; (*internal variable*)
		state : USINT; (*internal variable*)
		LockIDPar : USINT; (*internal variable*)
	END_VAR
END_FUNCTION_BLOCK

FUNCTION_BLOCK MC_DigitalCamSwitch (*allows a digital output (Track) to be set whenever the axis is inside a position window*)
	VAR_INPUT
		Axis : UDINT; (*axis reference*)
		Switches : MC_CAMSWITCH_REF; (*reference to the switching actions*)
		Outputs : MC_OUTPUT_REF; (*reference to the signal outputs*)
		TrackOptions : MC_TRACK_REF; (*reference to the track related properties*)
		Enable : BOOL; (*when set the FB parameters are downloaded*)
		EnableMask : UDINT; (*when set the digital outputs will be switched to ON and OFF*)
		InitSwitches : BOOL; (*initialize new switching action*)
		InitTrackOptions : BOOL; (*initialize new track related properties while switching is active*)
	END_VAR
	VAR_OUTPUT
		InOperation : BOOL; (*is set after all parameters have transferred*)
		Busy : BOOL; (*the function block is active*)
		SwitchesInitialized : BOOL; (*new switching actions initialized*)
		TrackOptionsInitialized : BOOL; (*new track related properties initialized*)
		Error : BOOL; (*error occurred in FB*)
		ErrorID : UINT; (*error number*)
	END_VAR
	VAR
		C_Master : UDINT; (*internal variable*)
		C_Slave : UDINT; (*internal variable*)
		C_Switches : MC_CAMSWITCH_REF; (*internal variable*)
		C_Outputs : MC_OUTPUT_REF; (*internal variable*)
		C_TrackOptions : MC_TRACK_REF; (*internal variable*)
		C_EnableMask : UDINT; (*internal variable*)
		C_CamConActRec : USINT; (*internal variable*)
		nextParRec : USINT; (*internal variable*)
		SelectRecMode : USINT; (*internal variable*)
		LockIDSend : USINT; (*internal variable*)
		C_InOperation : BOOL; (*internal variable*)
		C_Error : BOOL; (*internal variable*)
		C_ErrorID : UINT; (*internal variable*)
		C_Busy : BOOL; (*internal variable*)
		CC_ErrorID : UINT; (*internal variable*)
		EdgeInitSwitches : BOOL; (*internal variable*)
		EdgeInitTrackOptions : BOOL; (*internal variable*)
		CamConIndex : UINT; (*internal variable*)
		LogicIndex : UINT; (*internal variable*)
		VarIndex : UINT; (*internal variable*)
		CamConActRecOffset : UINT; (*internal variable*)
		CamConActRecRecIndex : USINT; (*internal variable*)
		LockIDMa : USINT; (*internal variable*)
		LockIDPar : USINT; (*internal variable*)
		LockID : USINT; (*internal variable*)
		sendSlot : USINT; (*internal variable*)
		readSlot : USINT; (*internal variable*)
		state : USINT; (*internal variable*)
		SptID : USINT; (*internal variable*)
		LockIDReceive : USINT; (*internal variable*)
	END_VAR
END_FUNCTION_BLOCK

FUNCTION_BLOCK MC_GearIn (*commands a ratio between the velocity of the master and slave axes*)
	VAR_INPUT
		Master : UDINT; (*axis reference of the master axis*)
		Slave : UDINT; (*axis reference of the slave axis*)
		Execute : BOOL; (*start the gearing process at the rising edge*)
		RatioNumerator : INT; (*gear ratio numerator*)
		RatioDenominator : UINT; (*gear ratio denominator*)
		Acceleration : REAL; (*maximum acceleration for gearing in*)
		Deceleration : REAL; (*maximum deceleration for gearing in*)
		MasterParID : UINT; (*use this master ParID instead of the set position*)
		MasterParIDMaxVelocity : REAL; (*maximum velocity of the master ParID*)
	END_VAR
	VAR_OUTPUT
		InGear : BOOL; (*commanded gearing complete*)
		Busy : BOOL; (*function block is not finished*)
		CommandAborted : BOOL; (*function block is aborted by another command*)
		Error : BOOL; (*error occurred in FB*)
		ErrorID : UINT; (*error number*)
	END_VAR
	VAR
		LockID : USINT; (*internal variable*)
		C_Master : UDINT; (*internal variable*)
		C_Slave : UDINT; (*internal variable*)
		C_Execute : BOOL; (*internal variable*)
		C_RatioNumerator : DINT; (*internal variable*)
		C_RatioDenominator : DINT; (*internal variable*)
		C_Acceleration : REAL; (*internal variable*)
		C_Deceleration : REAL; (*internal variable*)
		C_MasterParID : UINT; (*internal variable*)
		CC_ErrorID : UINT; (*internal variable*)
		C_MasterParIDMaxVelocity : REAL; (*internal variable*)
		C_InGear : BOOL; (*internal variable*)
		C_CommandAborted : BOOL; (*internal variable*)
		C_Error : BOOL; (*internal variable*)
		C_ErrorID : UINT; (*internal variable*)
		MpgenIndex : UINT; (*internal variable*)
		AutActualStateIndexOffset : UINT; (*internal variable*)
		AutActualStateIndexRecIndex : USINT; (*internal variable*)
		LockIDMa : USINT; (*internal variable*)
		sendSlot : USINT; (*internal variable*)
		readSlot : USINT; (*internal variable*)
		state : USINT; (*internal variable*)
		LockIDPar : USINT; (*internal variable*)
		MoveID : USINT; (*internal variable*)
		LockIDSend : USINT; (*internal variable*)
		LockIDReceive : USINT; (*internal variable*)
		SavedFrDrvCnt : USINT; (*internal variable*)
		WaitForTelegrams : BOOL; (*internal variable*)
	END_VAR
END_FUNCTION_BLOCK

FUNCTION_BLOCK MC_GearInPos (*commands a gear ratio between the position of the slave and master axis*)
	VAR_INPUT
		Master : UDINT; (*axis reference of the master axis*)
		Slave : UDINT; (*axis reference of the slave axis*)
		Execute : BOOL; (*start the gearing process at the rising edge*)
		RatioNumerator : INT; (*gear ration numerator*)
		RatioDenominator : UINT; (*gear ratio denominator*)
		MasterSyncPosition : REAL; (*master position at which the axes are running in sync*)
		SlaveSyncPosition : REAL; (*slave position at which the axes are running in sync*)
		SyncMode : USINT; (*defines the way to syncronize*)
		MasterStartDistance : REAL; (*master distance for preparation*)
		Velocity : REAL; (*maximum velocity during the time difference "StartSync" and "InSync"*)
		Acceleration : REAL; (*maximum acceleration during the time difference "StartSync" and "InSync"*)
		MasterParID : UINT; (*use this ParID from the master axis instead of the set position*)
		MasterParIDMaxVelocity : REAL; (*maximum value of the master ParID value*)
	END_VAR
	VAR_OUTPUT
		StartSync : BOOL; (*command gearing starts*)
		InSync : BOOL; (*commanded gearing is completed*)
		Busy : BOOL; (*function block is not finished*)
		CommandAborted : BOOL; (*function block is aborted by another command*)
		Error : BOOL; (*error occurred in FB*)
		ErrorID : UINT; (*error number*)
	END_VAR
	VAR
		C_Master : UDINT; (*internal variable*)
		C_Slave : UDINT; (*internal variable*)
		C_Execute : BOOL; (*internal variable*)
		C_RatioNumerator : DINT; (*internal variable*)
		C_RatioDenominator : DINT; (*internal variable*)
		Reserve1 : DINT; (*internal variable*)
		Reserve2 : DINT; (*internal variable*)
		C_SyncMode : USINT; (*internal variable*)
		LockID : USINT; (*internal variable*)
		LockIDPar : USINT; (*internal variable*)
		C_MasterStartDistance : DINT; (*internal variable*)
		C_MasterSyncPosition : DINT; (*internal variable*)
		C_SlaveSyncPosition : DINT; (*internal variable*)
		C_Velocity : REAL; (*internal variable*)
		C_Acceleration : REAL; (*internal variable*)
		C_MasterParID : UINT; (*internal variable*)
		C_MasterParIDMaxVelocity : REAL; (*internal variable*)
		C_StartSync : BOOL; (*internal variable*)
		C_InSync : BOOL; (*internal variable*)
		C_CommandAborted : BOOL; (*internal variable*)
		C_Error : BOOL; (*internal variable*)
		C_ErrorID : UINT; (*internal variable*)
		CC_Error : BOOL; (*internal variable*)
		MaPosition : DINT; (*internal variable*)
		DataTyp : UINT; (*internal variable*)
		MA_LastSyncPosition : DINT; (*internal variable*)
		SL_LastSyncPosition : DINT; (*internal variable*)
		MpgenIndex : UINT; (*internal variable*)
		Reserve3 : USINT; (*internal variable*)
		LockIDReceive : USINT; (*internal variable*)
		AutActualCamTypeOffset : UINT; (*internal variable*)
		AutActualCamTypeRecIndex : USINT; (*internal variable*)
		LockIDSend : USINT; (*internal variable*)
		AutActualStateIndexOffset : UINT; (*internal variable*)
		AutActualStateIndexRecIndex : USINT; (*internal variable*)
		LockIDMa : USINT; (*internal variable*)
		sendSlot : USINT; (*internal variable*)
		readSlot : USINT; (*internal variable*)
		state : USINT; (*internal variable*)
		MoveID : USINT; (*internal variable*)
		CC_ErrorID : UINT; (*internal variable*)
		Reserve4 : UINT; (*internal variable*)
	END_VAR
END_FUNCTION_BLOCK

FUNCTION_BLOCK MC_GearOut (*disengages the geared slave from the master axis*)
	VAR_INPUT
		Slave : UDINT; (*axis reference of slave axis*)
		Execute : BOOL; (*start disengaging process at rising edge*)
	END_VAR
	VAR_OUTPUT
		Done : BOOL; (*disengaging completed*)
		Busy : BOOL; (*function block is not finished*)
		Error : BOOL; (*error occurred in FB*)
		ErrorID : UINT; (*error number*)
	END_VAR
	VAR
		C_Slave : UDINT; (*internal variable*)
		C_Execute : BOOL; (*internal variable*)
		C_Done : BOOL; (*internal variable*)
		C_Error : BOOL; (*internal variable*)
		C_ErrorID : UINT; (*internal variable*)
		state : USINT; (*internal variable*)
		LockIDPar : USINT; (*internal variable*)
		MoveID : USINT; (*internal variable*)
	END_VAR
END_FUNCTION_BLOCK

FUNCTION_BLOCK MC_Halt (*commands a controlled motion stop*)
	VAR_INPUT
		Axis : UDINT; (*axis reference*)
		Execute : BOOL; (*start the action at rising edge*)
		Deceleration : REAL; (*value of deceleration*)
	END_VAR
	VAR_OUTPUT
		Done : BOOL; (*zero velocity is reached*)
		Busy : BOOL; (*function block is not finished*)
		CommandAborted : BOOL; (*function block aborted by calling another movement function block*)
		Error : BOOL; (*error occurred in FB*)
		ErrorID : UINT; (*error number*)
	END_VAR
	VAR
		C_Axis : UDINT; (*internal variable*)
		C_Execute : BOOL; (*internal variable*)
		cmdExecute : BOOL; (*internal variable*)
		C_Done : BOOL; (*internal variable*)
        C_CommandAborted : BOOL; (*internal variable*)
        C_Deceleration : REAL; (*internal variable*)
		C_ErrorID : UINT; (*internal variable*)
		C_Error : BOOL; (*internal variable*)
		state : USINT; (*internal variable*)
		MoveID : USINT; (*internal variable*)
        LockIDPar : USINT; (*internal variable*)
        Reserve : UINT; (*internal variable*)
	END_VAR
END_FUNCTION_BLOCK

FUNCTION_BLOCK MC_Home (*starts the homing movement of an axis according to the homing parameters*)
	VAR_INPUT
		Axis : UDINT; (*axis reference*)
		Execute : BOOL; (*start movement at rising edge*)
		Position : REAL; (*absolute position when the reference signal is detected*)
		HomingMode : USINT; (*select the homing mode*)
	END_VAR
	VAR_OUTPUT
		Done : BOOL; (*homing procedure has finished successfully*)
		Busy : BOOL; (*function block is not finished*)
		CommandAborted : BOOL; (*function block is aborted by another command*)
		Error : BOOL; (*error occurred in FB*)
		ErrorID : UINT; (*error number*)
	END_VAR
	VAR
		C_Axis : UDINT; (*internal variable*)
		C_Execute : BOOL; (*internal variable*)
		C_Position : DINT; (*internal variable*)
		C_HomingMode : USINT; (*internal variable*)
		LockIDPar : USINT; (*internal variable*)
		C_Done : BOOL; (*internal variable*)
		C_CommandAborted : BOOL; (*internal variable*)
		C_Error : BOOL; (*internal variable*)
		C_ErrorID : UINT; (*internal variable*)
		state : USINT; (*internal variable*)
		MoveID : USINT; (*internal variable*)
		CC_Position : REAL; (*internal variable*)
	END_VAR
END_FUNCTION_BLOCK

FUNCTION_BLOCK MC_LimitLoad (*limits the motor torque to a set value*)
	VAR_INPUT
		Axis : UDINT; (*axis reference*)
		Enable : BOOL; (*when set limitation is activated*)
		Load : REAL; (*limit value for the motor torque [Nm]*)
		Direction : USINT; (*movement direction*)
	END_VAR
	VAR_OUTPUT
		Busy : BOOL; (*function block is not finished*)
		Ready : BOOL; (*parameters initialized*)
		Active : BOOL; (*torque is limited*)
		Error : BOOL; (*error occurred in FB*)
		ErrorID : UINT; (*error number*)
	END_VAR
	VAR
		C_Axis : UDINT; (*internal variable*)
		IS : MC_0133_IS_TYP; (*internal variable*)
	END_VAR
END_FUNCTION_BLOCK

FUNCTION_BLOCK MC_MoveAbsolute (*commands a controlled motion at a specified absolute position*)
	VAR_INPUT
		Axis : UDINT; (*axis reference*)
		Execute : BOOL; (*start movement at rising edge*)
		Position : REAL; (*target position for the motion*)
		Velocity : REAL; (*maximum velocity*)
		Acceleration : REAL; (*maximum acceleration*)
		Deceleration : REAL; (*maximum deceleration*)
		Direction : USINT; (*movement direction*)
	END_VAR
	VAR_OUTPUT
		Done : BOOL; (*commanded position reached*)
		Busy : BOOL; (*function block is not finished*)
		CommandAborted : BOOL; (*function block aborted by another command*)
		Error : BOOL; (*error occurred in FB*)
		ErrorID : UINT; (*error number*)
	END_VAR
	VAR
		C_Axis : UDINT; (*internal variable*)
		C_Execute : BOOL; (*internal variable*)
		cmdExecute : BOOL; (*internal variable*)
        C_Direction : USINT; (*internal variable*)
        LockIDPar : USINT; (*internal variable*)
        C_Position : DINT; (*internal variable*)
        C_Velocity : REAL; (*internal variable*)
        C_Acceleration : REAL; (*internal variable*)
        C_Deceleration : REAL; (*internal variable*)
        C_Done : BOOL; (*internal variable*)
		C_CommandAborted : BOOL; (*internal variable*)
        C_Error : BOOL; (*internal variable*)
        state : USINT; (*internal variable*)
        C_CommandedOffset : DINT; (*internal variable*)
		C_ErrorID : UINT; (*internal variable*)
        MoveID : USINT; (*internal variable*)
        oldMoveID : USINT; (*internal variable*)
	END_VAR
END_FUNCTION_BLOCK

FUNCTION_BLOCK MC_MoveAdditive (*commands a controlled motion of a specified relative distance*)
	VAR_INPUT
		Axis : UDINT; (*axis reference*)
		Execute : BOOL; (*start movement at rising edge*)
		Distance : REAL; (*relative distance for the motion*)
		Velocity : REAL; (*maximum velocity for the motion*)
		Acceleration : REAL; (*maximum acceleration for the motion*)
		Deceleration : REAL; (*maximum deceleration for the motion*)
	END_VAR
	VAR_OUTPUT
		Done : BOOL; (*commanded position reached*)
		Busy : BOOL; (*function block is not finished*)
		CommandAborted : BOOL; (*function block aborted by another command*)
		Error : BOOL; (*error occurred in FB*)
		ErrorID : UINT; (*error number*)
	END_VAR
	VAR
		C_Axis : UDINT; (*internal variable*)
		C_Distance : DINT; (*internal variable*)
		C_Velocity : REAL; (*internal variable*)
		C_Acceleration : REAL; (*internal variable*)
        C_Deceleration : REAL; (*internal variable*)
        C_Execute : BOOL; (*internal variable*)
		cmdExecute : BOOL; (*internal variable*)
		C_Done : BOOL; (*internal variable*)
		C_CommandAborted : BOOL; (*internal variable*)
		C_CommandedPosition : DINT; (*internal variable*)
        C_CommandedOffset : DINT; (*internal variable*)
        C_ErrorID : UINT; (*internal variable*)
        C_Error : BOOL; (*internal variable*)
		state : USINT; (*internal variable*)
		LockIDPar : USINT; (*internal variable*)
        MoveID : USINT; (*internal variable*)
        oldMoveID : USINT; (*internal variable*)
        Reserve : USINT; (*internal variable*)
	END_VAR
END_FUNCTION_BLOCK

FUNCTION_BLOCK MC_MoveVelocity (*commands a motion with specified velocity*)
	VAR_INPUT
		Axis : UDINT; (*axis reference*)
		Execute : BOOL; (*start movement at rising edge*)
		Velocity : REAL; (*Value of maximum velocity*)
		Acceleration : REAL; (*Value of maximum acceleration*)
		Deceleration : REAL; (*Value of maximum deceleration*)
		Direction : USINT; (*direction of movement*)
	END_VAR
	VAR_OUTPUT
		InVelocity : BOOL; (*commanded velocity reached*)
		Busy : BOOL; (*function block is not finished*)
		CommandAborted : BOOL; (*function block aborted by another command*)
		Error : BOOL; (*error occurred in FB*)
		ErrorID : UINT; (*error number*)
	END_VAR
	VAR
		C_Axis : UDINT; (*internal variable*)
		C_Execute : BOOL; (*internal variable*)
		cmdExecute : BOOL; (*internal variable*)
		C_Velocity : REAL; (*internal variable*)
		C_Acceleration : REAL; (*internal variable*)
		C_Deceleration : REAL; (*internal variable*)
		C_Direction : USINT; (*internal variable*)
		LockIDPar : USINT; (*internal variable*)
		C_InVelocity : BOOL; (*internal variable*)
		C_CommandAborted : BOOL; (*internal variable*)
		C_Error : BOOL; (*internal variable*)
		C_ErrorID : UINT; (*internal variable*)
		state : USINT; (*internal variable*)
		MoveID : USINT; (*internal variable*)
	END_VAR
END_FUNCTION_BLOCK

FUNCTION_BLOCK MC_Phasing (*creates a phase shift in the master position of a slave axis*)
	VAR_INPUT
		Master : UDINT; (*axis reference of the master axis*)
		Slave : UDINT; (*axis reference of the slave axis*)
		Execute : BOOL; (*start the phasing process at rising edge*)
		PhaseShift : REAL; (*phase difference*)
		Velocity : REAL; (*maximum velocity to reach phase difference*)
		Acceleration : REAL; (*maximum acceleration to reach phase difference*)
	END_VAR
	VAR_OUTPUT
		Done : BOOL; (*commanded phasing reached*)
		Busy : BOOL; (*function block is not finished*)
		CommandAborted : BOOL; (*function block aborted by another command*)
		Error : BOOL; (*error occurred in FB*)
		ErrorID : UINT; (*error number*)
	END_VAR
	VAR
		C_Master : UDINT; (*internal variable*)
		C_Slave : UDINT; (*internal variable*)
		C_Execute : BOOL; (*internal variable*)
		C_PhaseShift : DINT; (*internal variable*)
		C_Velocity : REAL; (*internal variable*)
		C_Acceleration : REAL; (*internal variable*)
		C_Done : BOOL; (*internal variable*)
		C_CommandAborted : BOOL; (*internal variable*)
		C_Error : BOOL; (*internal variable*)
		C_ErrorID : UINT; (*internal variable*)
		MpgenIndex : UINT; (*internal variable*)
		MpgenStatusOffset : UINT; (*internal variable*)
		MpgenStatusRecIndex : USINT; (*internal variable*)
		LockIDPar : USINT; (*internal variable*)
		SavedFrDrvCnt : USINT; (*internal variable*)
		state : USINT; (*internal variable*)
		FbID : USINT; (*internal variable*)
		WaitForTelegrams : BOOL; (*internal variable*)
	END_VAR
END_FUNCTION_BLOCK

FUNCTION_BLOCK MC_Power (*switches on the controller of the axis*)
	VAR_INPUT
		Axis : UDINT; (*axis reference*)
		Enable : BOOL; (*as long as "Enable" is TRUE, the drive power stage is enabled*)
	END_VAR
	VAR_OUTPUT
		Status : BOOL; (*effective status of the power stage*)
		Busy : BOOL; (*function block is not finished*)
		Error : BOOL; (*error occurred in FB*)
		ErrorID : UINT; (*error number*)
	END_VAR
	VAR
		state : USINT; (*internal variable*)
		C_Error : BOOL; (*internal variable*)
		C_ErrorID : UINT; (*internal variable*)
		C_Axis : UDINT; (*internal variable*)
		startTicks : UDINT; (*internal variable*)
		AxisTypeCtrlOffAxisState : UINT; (*internal variable*)
	END_VAR
END_FUNCTION_BLOCK

FUNCTION_BLOCK MC_ReadActualPosition (*returns the actual axis position*)
	VAR_INPUT
		Axis : UDINT; (*axis reference*)
		Enable : BOOL; (*when set the position is read*)
	END_VAR
	VAR_OUTPUT
		Valid : BOOL; (*output of FB is valid*)
		Busy : BOOL; (*the function block is not finished*)
		Error : BOOL; (*error occurred in FB*)
		ErrorID : UINT; (*error number*)
		Position : REAL; (*actual position of the axis*)
	END_VAR
	VAR
		C_Axis : UDINT; (*internal variable*)
		C_ErrorID : UINT; (*internal variable*)
		C_Error : BOOL; (*internal variable*)
		state : USINT; (*internal variable*)
	END_VAR
END_FUNCTION_BLOCK

FUNCTION_BLOCK MC_ReadActualTorque (*returns the axis torque*)
	VAR_INPUT
		Axis : UDINT; (*axis reference*)
		Enable : BOOL; (*read the actual torque continuously while enabled*)
	END_VAR
	VAR_OUTPUT
		Valid : BOOL; (*output is available*)
		Busy : BOOL; (*function block is not finished*)
		Error : BOOL; (*error occurred in FB*)
		ErrorID : UINT; (*error number*)
		Torque : REAL; (*value of the actual torque*)
	END_VAR
	VAR
		C_Axis : UDINT; (*internal variable*)
		TorqueOffset : UINT; (*internal variable*)
		TorqueRecIndex : USINT; (*internal variable*)
		LockID : USINT; (*internal variable*)
		C_ErrorID : UINT; (*internal variable*)
		C_Error : BOOL; (*internal variable*)
		state : USINT; (*internal variable*)
		LockIDPar : USINT; (*internal variable*)
	END_VAR
END_FUNCTION_BLOCK

FUNCTION_BLOCK MC_ReadActualVelocity (*returns the axis velocity*)
	VAR_INPUT
		Axis : UDINT; (*axis reference*)
		Enable : BOOL; (*read the velocity continuously while enabled*)
	END_VAR
	VAR_OUTPUT
		Valid : BOOL; (*output is available*)
		Busy : BOOL; (*function block is not finished*)
		Error : BOOL; (*error occurred in FB*)
		ErrorID : UINT; (*error number*)
		Velocity : REAL; (*value of actual velocity*)
	END_VAR
	VAR
		C_Axis : UDINT; (*internal variable*)
		C_ErrorID : UINT; (*internal variable*)
		C_Error : BOOL; (*internal variable*)
		state : USINT; (*internal variable*)
	END_VAR
END_FUNCTION_BLOCK

FUNCTION_BLOCK MC_ReadAxisError (*returns the actual axis error as long as "Enable" is TRUE*)
	VAR_INPUT
		Axis : UDINT; (*axis reference*)
		Enable : BOOL; (*read error number/text*)
		Acknowledge : BOOL; (*acknowledge current axis error*)
		DataAddress : UDINT; (*address of error text string*)
		DataLength : UINT; (*length of error text string*)
		DataObjectName : STRING[12]; (*name of error text module*)
	END_VAR
	VAR_OUTPUT
		Valid : BOOL; (*error text is valid*)
		Busy : BOOL; (*function block is not finished*)
		Error : BOOL; (*error occurred in FB*)
		ErrorID : UINT; (*error number*)
		AxisErrorID : UINT; (*axis error number*)
		AxisErrorCount : UINT; (*count of axis error*)
	END_VAR
	VAR
		C_Axis : UDINT; (*internal variable*)
		C_Acknowledge : BOOL; (*internal variable*)
		C_OldAcknowledge : BOOL; (*internal variable*)
		C_DataObjectName : STRING[12]; (*internal variable*)
		Reserve : UINT; (*internal variable*)
		writeText : BOOL; (*internal variable*)
		C_Error : BOOL; (*internal variable*)
		C_ErrorID : UINT; (*internal variable*)
		state : USINT; (*internal variable*)
	END_VAR
END_FUNCTION_BLOCK

FUNCTION_BLOCK MC_ReadBoolParameter (*returns the value of one Boolean PLCopen parameter*)
	VAR_INPUT
		Axis : UDINT; (*axis reference*)
		Enable : BOOL; (*get the value of the parameter while enabled*)
		ParameterNumber : INT; (*number of the parameter*)
	END_VAR
	VAR_OUTPUT
		Valid : BOOL; (*parameter available*)
		Busy : BOOL; (*function block is not finished*)
		Error : BOOL; (*error occurred in FB*)
		ErrorID : UINT; (*error number*)
		Value : BOOL; (*value of requested parameter*)
	END_VAR
	VAR
		C_Axis : UDINT; (*internal variable*)
		C_ErrorID : UINT; (*internal variable*)
		C_Error : BOOL; (*internal variable*)
		state : USINT; (*internal variable*)
	END_VAR
END_FUNCTION_BLOCK

FUNCTION_BLOCK MC_ReadDigitalInput (*reads an digital input on an ACOPOS plug-in module*)
	VAR_INPUT
		Input : MC_INPUT_REF; (*reference to input signal source*)
		Enable : BOOL; (*get value of selected input signal continuously while enabled*)
	END_VAR
	VAR_OUTPUT
		Valid : BOOL; (*input signal value is valid*)
		Busy : BOOL; (*function block is not finished*)
		Error : BOOL; (*error occurred in FB*)
		ErrorID : UINT; (*error number*)
		Value : BOOL; (*value of selected input signal*)
	END_VAR
	VAR
		C_Axis : UDINT; (*internal variable*)
		C_Input : MC_INPUT_REF; (*internal variable*)
		C_Error : BOOL; (*internal variable*)
		C_ErrorID : UINT; (*internal variable*)
		ReadDigitalInputOffset : UINT; (*internal variable*)
		ReadDigitalInputRecIndex : USINT; (*internal variable*)
		LockID : USINT; (*internal variable*)
		ReadDigitalInputValue : UINT; (*internal variable*)
		ReadDigitalInputMask : UINT; (*internal variable*)
		state : USINT; (*internal variable*)
		LockIDPar : USINT; (*internal variable*)
	END_VAR
END_FUNCTION_BLOCK

FUNCTION_BLOCK MC_ReadDigitalOutput (*reads a digital output*)
	VAR_INPUT
		Output : MC_OUTPUT_REF; (*reference to signal outputs*)
		Enable : BOOL; (*get value of selected output signal continouosly while enabled*)
	END_VAR
	VAR_OUTPUT
		Valid : BOOL; (*output signal value is valid*)
		Busy : BOOL; (*function block is not finished*)
		Error : BOOL; (*error occurred in FB*)
		ErrorID : UINT; (*error number*)
		Value : BOOL; (*value of selected output signal*)
	END_VAR
	VAR
		C_Axis : UDINT; (*internal variable*)
		C_Output : MC_OUTPUT_REF; (*internal variable*)
		C_Error : BOOL; (*internal variable*)
		C_ErrorID : UINT; (*internal variable*)
		ReadDigitalOutputOffset : UINT; (*internal variable*)
		ReadDigitalOutputRecIndex : USINT; (*internal variable*)
		LockID : USINT; (*internal variable*)
		ReadDigitalOutputValue : UINT; (*internal variable*)
		ReadDigitalOutputMask : UINT; (*internal variable*)
		state : USINT; (*internal variable*)
		LockIDPar : USINT; (*internal variable*)
	END_VAR
END_FUNCTION_BLOCK

FUNCTION_BLOCK MC_ReadParameter (*returns the value of a specific PLCopen parameter*)
	VAR_INPUT
		Axis : UDINT; (*axis reference*)
		Enable : BOOL; (*get the value of the parameter while enabled*)
		ParameterNumber : INT; (*number of parameter*)
	END_VAR
	VAR_OUTPUT
		Valid : BOOL; (*parameter available*)
		Busy : BOOL; (*function block is not finished*)
		Error : BOOL; (*error occurred in FB*)
		ErrorID : UINT; (*error number*)
		Value : REAL; (*value of the requested parameter*)
	END_VAR
	VAR
		C_Axis : UDINT; (*internal variable*)
		C_ErrorID : UINT; (*internal variable*)
		C_Error : BOOL; (*internal variable*)
		state : USINT; (*internal variable*)
		LockIDPar : USINT; (*internal variable*)
	END_VAR
END_FUNCTION_BLOCK

FUNCTION_BLOCK MC_ReadStatus (*returns the detailed status of the motion currently in progress*)
	VAR_INPUT
		Axis : UDINT; (*axis reference*)
		Enable : BOOL; (*read the axis status continuously while enabled*)
	END_VAR
	VAR_OUTPUT
		Valid : BOOL; (*true if valid outputs available*)
		Busy : BOOL; (*the function block is not finished*)
		Error : BOOL; (*error occurred in FB*)
		ErrorID : UINT; (*error number*)
		Errorstop : BOOL; (*an error occurred on the drive*)
		Disabled : BOOL; (*controller is switched off*)
		Stopping : BOOL; (*MC_Stop is active*)
		StandStill : BOOL; (*controller is switched on but no motion is active*)
		DiscreteMotion : BOOL; (*axis executes an absolute or an additive motion*)
		ContinuousMotion : BOOL; (*axis is in permanent motion*)
		SynchronizedMotion : BOOL; (*axis is synchronized with another axis*)
		Homing : BOOL; (*MC_Home has started homing the axis*)
	END_VAR
	VAR
		C_Axis : UDINT; (*internal variable*)
		C_Error : BOOL; (*internal variable*)
		C_ErrorID : UINT; (*internal variable*)
		state : USINT; (*internal variable*)
	END_VAR
END_FUNCTION_BLOCK

FUNCTION_BLOCK MC_Reset (*makes transition from Errorstop to Standstill or Disabled by resetting internal axis related errors*)
	VAR_INPUT
		Axis : UDINT; (*axis reference*)
		Execute : BOOL; (*resets the axis at the rising edge*)
	END_VAR
	VAR_OUTPUT
		Done : BOOL; (*standstill state is reached*)
		Busy : BOOL; (*function block is not finished*)
		Error : BOOL; (*error occurred in FB*)
		ErrorID : UINT; (*error number*)
	END_VAR
	VAR
		C_Axis : UDINT; (*internal variable*)
		C_ErrorID : UINT; (*internal variable*)
		C_Error : BOOL; (*internal variable*)
		state : USINT; (*internal variable*)
	END_VAR
END_FUNCTION_BLOCK

FUNCTION_BLOCK MC_SetOverride (*sets the values of override parameters for velocity and acceleration/deceleration*)
	VAR_INPUT
		Axis : UDINT; (*axis reference*)
		Enable : BOOL; (*write the value of the override at the rising edge*)
		VelFactor : REAL; (*new override factor for the velocity*)
		AccFactor : REAL; (*new override factor for the acceleration/deceleration*)
	END_VAR
	VAR_OUTPUT
		Enabled : BOOL; (*override successfully written*)
		Busy : BOOL; (*function block not finished*)
		Error : BOOL; (*error occurred in FB*)
		ErrorID : UINT; (*error number*)
	END_VAR
	VAR
		C_Axis : UDINT; (*internal variable*)
		C_VelFactor : REAL; (*internal variable*)
		C_AccFactor : REAL; (*internal variable*)
		OldVelFactor : REAL; (*internal variable*)
		C_ErrorID : UINT; (*internal variable*)
		C_Error : BOOL; (*internal variable*)
		state : USINT; (*internal variable*)
	END_VAR
END_FUNCTION_BLOCK

FUNCTION_BLOCK MC_Stop (*commands a controlled motion stop and transfers the axis to the state Stopping*)
	VAR_INPUT
		Axis : UDINT; (*axis reference*)
		Execute : BOOL; (*start the action at rising edge*)
		Deceleration : REAL; (*value of deceleration *)
	END_VAR
	VAR_OUTPUT
		Done : BOOL; (*zero velocity is reached*)
		Busy : BOOL; (*function block is not finished*)
		CommandAborted : BOOL; (*function block is aborted by switching off power*)
		Error : BOOL; (*error occurred in FB*)
		ErrorID : UINT; (*error number*)
	END_VAR
	VAR
		C_Axis : UDINT; (*internal variable*)
		C_Execute : BOOL; (*internal variable*)
		C_Error : BOOL; (*internal variable*)
		C_ErrorID : UINT; (*internal variable*)
		C_Deceleration : REAL; (*internal variable*)
		C_CommandAborted : BOOL; (*internal variable*)
		state : USINT; (*internal variable*)
		MoveID : USINT; (*internal variable*)
	END_VAR
END_FUNCTION_BLOCK

FUNCTION_BLOCK MC_TouchProbe (*records an axis position at a trigger event*)
	VAR_INPUT
		Axis : UDINT; (*axis reference*)
		TriggerInput : MC_TRIGGER_REF; (*trigger input signal source*)
		Execute : BOOL; (*transfer parameters at rising edge*)
		WindowOnly : BOOL; (*if set, only use the window to accept trigger events*)
		FirstPosition : REAL; (*start position from where trigger events are accepted*)
		LastPosition : REAL; (*end position of the window*)
	END_VAR
	VAR_OUTPUT
		Done : BOOL; (*trigger event recorded*)
		Busy : BOOL; (*function block not finished*)
		CommandAborted : BOOL; (*function block is aborted by another command*)
		Error : BOOL; (*error occurred in FB*)
		ErrorID : UINT; (*error number*)
		RecordedPosition : REAL; (*position where the trigger event occurred*)
	END_VAR
	VAR
		C_Axis : UDINT; (*internal variable*)
		C_Done : BOOL; (*internal variable*)
		C_Busy : BOOL; (*internal variable*)
		C_TriggerInput : MC_TRIGGER_REF; (*internal variable*)
		C_Execute : BOOL; (*internal variable*)
		C_WindowOnly : BOOL; (*internal variable*)
		C_FirstPosition : DINT; (*internal variable*)
		C_LastPosition : DINT; (*internal variable*)
		C_Error : BOOL; (*internal variable*)
		C_ErrorID : UINT; (*internal variable*)
		C_CommandAborted : BOOL; (*internal variable*)
		C_RecordedPosition : DINT; (*internal variable*)
		InputSourceChanged : BOOL; (*internal variable*)
		EdgeChanged : BOOL; (*internal variable*)
		PosSourceChanged : BOOL; (*internal variable*)
		SavedToDrvCnt : USINT; (*internal variable*)
		Reserve2 : USINT; (*internal variable*)
		state : USINT; (*internal variable*)
		LockID : USINT; (*internal variable*)
		LockIDPar : USINT; (*internal variable*)
		cycleTime : UINT; (*internal variable*)
		LatchPos : DINT; (*internal variable*)
		LatchStatusOffset : UINT; (*internal variable*)
		LatchStatusRecIndex : USINT; (*internal variable*)
		Reserve1 : USINT; (*internal variable*)
		LatchPosOffset : UINT; (*internal variable*)
		LatchPosRecIndex : USINT; (*internal variable*)
		SptID : USINT; (*internal variable*)
	END_VAR
END_FUNCTION_BLOCK

FUNCTION_BLOCK MC_TorqueControl (*starts a torque movement with limited speed*)
	VAR_INPUT
		Axis : UDINT; (*axis reference*)
		Execute : BOOL; (*start movement at rising edge*)
		Torque : REAL; (*signed set torque value for the axis [Nm]*)
		TorqueRamp : REAL; (*torque increase while reaching "Torque" [Nm/s]*)
		Velocity : REAL; (*velocity limit for axis*)
		Acceleration : REAL; (*maximum acceleration or deceleration*)
	END_VAR
	VAR_OUTPUT
		InTorque : BOOL; (*set torque value reached*)
		Busy : BOOL; (*function block is not finished*)
		Active : BOOL; (*function block is controlling the axis*)
		CommandAborted : BOOL; (*command is aborted by another command*)
		Error : BOOL; (*error occured in FB*)
		ErrorID : UINT; (*error number*)
		AxisLimitActive : BOOL; (*axis velocity limited*)
	END_VAR
	VAR
		C_Axis : UDINT; (*internal variable*)
		IS : MC_0096_IS_TYP; (*internal variable*)
	END_VAR
END_FUNCTION_BLOCK

FUNCTION_BLOCK MC_BR_TorqueControl (*starts a torque movement with limited speed*)
	VAR_INPUT
		Axis : UDINT; (*axis reference*)
		Enable : BOOL; (*function block is activated*)
		InitData : BOOL; (*parameter change while the FB is active*)
		StartSignal : BOOL; (*starts torque-controlled movement*)
		Torque : REAL; (*signed set torque value for the axis [Nm]*)
		TorqueRamp : REAL; (*torque increase while reaching "Torque" [Nm/s]*)
		PosMaxVelocity : REAL; (*velocity limit for axis*)
		NegMaxVelocity : REAL; (*velocity limit for axis*)
		Acceleration : REAL; (*maximum acceleration or deceleration*)
		Mode : UINT; (*mode selection (bit coded)*)
		TimeLimit : REAL; (*maximum movement time with limited speed or acceleration*)
		StartParID : UINT; (*not used at the moment*)
		TorqueParID : UINT; (*set torque value from ParID*)
	END_VAR
	VAR_OUTPUT
		InTorque : BOOL; (*set torque reached*)
		Busy : BOOL; (*function block is not finished*)
		Active : BOOL; (*function block is controlling the axis*)
		CommandAborted : BOOL; (*command is aborted by another command*)
		Error : BOOL; (*error occured in FB*)
		ErrorID : UINT; (*error number*)
		DataInitialized : BOOL; (*parameter online change done*)
		WaitingForStart : BOOL; (*ready for start via "StartSignal"*)
		AxisLimitActive : BOOL; (*axis velocity or acceleration limited*)
	END_VAR
	VAR
		C_Axis : UDINT; (*internal variable*)
		IS : MC_0100_IS_TYP; (*internal variable*)
	END_VAR
END_FUNCTION_BLOCK

FUNCTION_BLOCK MC_WriteBoolParameter (*writes the value of one Boolean PLCopen parameter*)
	VAR_INPUT
		Axis : UDINT; (*axis reference*)
		Execute : BOOL; (*write the value of the parameter at rising edge*)
		ParameterNumber : INT; (*number of the parameter*)
		Value : BOOL; (*new value of specified parameter*)
	END_VAR
	VAR_OUTPUT
		Done : BOOL; (*parameter successfully written*)
		Busy : BOOL; (*function block is not finished*)
		Error : BOOL; (*error occurred in FB*)
		ErrorID : UINT; (*error number*)
	END_VAR
	VAR
		C_Axis : UDINT; (*internal variable*)
		C_ParameterNumber : INT; (*internal variable*)
		Reserve : UINT; (*internal variable*)
		state : USINT; (*internal variable*)
	END_VAR
END_FUNCTION_BLOCK

FUNCTION_BLOCK MC_WriteDigitalOutput (*writes a digital output*)
	VAR_INPUT
		Output : MC_OUTPUT_REF; (*reference to signal output*)
		Execute : BOOL; (*write the value of selected output*)
		Value : BOOL; (*the value of the selected output*)
	END_VAR
	VAR_OUTPUT
		Done : BOOL; (*writing of the output signal value is done*)
		Busy : BOOL; (*function block is not finished*)
		Error : BOOL; (*error occurred in FB*)
		ErrorID : UINT; (*error number*)
	END_VAR
	VAR
		C_Axis : UDINT; (*internal variable*)
		C_Output : MC_OUTPUT_REF; (*internal variable*)
		C_Execute : BOOL; (*internal variable*)
		C_Value : BOOL; (*internal variable*)
		C_Done : BOOL; (*internal variable*)
		C_Error : BOOL; (*internal variable*)
		C_ErrorID : UINT; (*internal variable*)
		WriteDigitalOutputMask : UINT; (*internal variable*)
		state : USINT; (*internal variable*)
		LockIDPar : USINT; (*internal variable*)
	END_VAR
END_FUNCTION_BLOCK

FUNCTION_BLOCK MC_WriteParameter (*writes the value to a specific PLCopen parameter*)
	VAR_INPUT
		Axis : UDINT; (*axis reference*)
		Execute : BOOL; (*write the value of the parameter at the rising edge*)
		ParameterNumber : INT; (*number of the parameter*)
		Value : REAL; (*new value of specified parameter*)
	END_VAR
	VAR_OUTPUT
		Done : BOOL; (*parameter succesfully written*)
		Busy : BOOL; (*function block is not finished*)
		Error : BOOL; (*error occurred in FB*)
		ErrorID : UINT; (*error number*)
	END_VAR
	VAR
		C_Axis : UDINT; (*internal variable*)
		C_Execute : BOOL; (*internal variable*)
		C_ParameterNumber : INT; (*internal variable*)
		C_Value : REAL; (*internal variable*)
		C_Done : BOOL; (*internal variable*)
		C_Error : BOOL; (*internal variable*)
		C_ErrorID : UINT; (*internal variable*)
		state : USINT; (*internal variable*)
		LockIDPar : USINT; (*internal variable*)
	END_VAR
END_FUNCTION_BLOCK

(* ---- acp10_mc.var ---- *)
VAR CONSTANT
	mc5TH_ORDER_POLYNOMIAL : UINT := 4; (*motion rule*)
	mcABOVE_WINDOW : USINT := 40; (*trigger event mode*)
	mcABS : USINT := 1; (*encoder type*)
	mcABSOLUTE : USINT := 0; (*start mode*)
	mcABSOLUTE_NO_RESET : USINT := 2; (*definition for the shift input of MC_BR_Offset and MC_BR_Phasing*)
	mcACKNOWLEDGE_ALL : UINT := 2; (*acknowledge all error records immediately*)
	mcACT_CFG : UINT := 1;
	mcACTUAL_POSITION : UINT := 1; (*position source for MPDC*)
	mcACTUAL_VELOCITY : INT := 10; (*PLCopen motion parameter*)
	mcADD_DATE_TIME : UINT := 1; (*additional data object type*)
	mcALL_AXES : UDINT := 16#FFFFFFFF;
	mcALL_EVENTS : USINT := 255; (*event index*)
	mcALL_PARAMS : USINT := 0; (*parameter index*)
	mcALL_STATES : USINT := 255; (*state index*)
	mcAUT_POS_TOLERANCE : INT := 1009; (*PLCopen motion parameter*)
	mcAUTOMAT_POS : USINT := 100; (*additional movement direction*)
	mcAVERAGE : UINT := 2;
	mcAVERAGE_WEIGHTED : UINT := 4;
	mcAXIS_ERROR : USINT := 0;
	mcAXIS_FACTOR : INT := 1007; (*PLCopen motion parameter*)
	mcAXIS_FACTOR_MAPPING : INT := 1019; (*PLCopen motion parameter*)
	mcAXIS_NETWORK_CYCLE_TIME: INT := 1018; (*PLCopen motion parameter*)
	mcAXIS_PERIOD : INT := 1008; (*PLCopen motion parameter*)
	mcAXIS_PERIOD_MAPPING : INT := 1020; (*PLCopen motion parameter*)
	mcAXIS_WARNING : USINT := 1;
	mcBASIS_PARAMETERS : REAL := 2.0; (*Option for DefaultMoveParameter*)
	mcBELOW_WINDOW : USINT := 50; (*trigger event mode*)
	mcBESTFIT_5TH_ORDER : UINT := 1024; (*interpolation rule*)
	mcBESTFIT_6TH_ORDER : UINT := 1280; (*interpolation rule*)
	mcBLANK : UINT := 0;
	mcBRAKE_CONTROL_INIT : USINT := 8; (*brake command*)
	mcBRAKE_TEST_INIT : USINT := 2; (*brake command*)
	mcBRAKE_TEST_START : USINT := 4; (*brake command*)
	mcCALCULATION : UINT := 11; (*setup mode*)
	mcCATCH_UP : USINT := 4; (*synchronization mode*)
	mcCHECK : UINT := 1; (*mode for automat compensation check*)
	mcCHECK_HOMING_OFF : USINT := 1; (*disable homing check*)
	mcCLOSE : USINT := 0;
	mcCMD_ERROR : UINT := 1; (*error command*)
    mcCMD_ERROR_COAST_TO_STANDSTILL : UINT := 5; (*error command*)
    mcCMD_ERROR_INDUCTION_HALT : UINT := 6; (*error command*)
	mcCMD_ERROR_STOP : UINT := 2; (*error command*)
	mcCMD_ERROR_STOP_CTRL_OFF : UINT := 3; (*error command*)
	mcCMD_ERROR_V_STOP_CTRL_OFF : UINT := 4; (*error command*)
	mcCMD_WARNING : UINT := 0; (*error command *)
	mcCOMMANDED_POSITION : INT := 1; (*PLCopen motion parameter*)
	mcCOMMANDED_VELOCITY : INT := 11; (*PLCopen motion parameter*)
	mcCONTINUE_CONTROLLER_OFF : UINT := 128; (* continue if controller is off *)
	mcCORRECT_CURRENT_CYCLE : UINT := 32768; (*additive StartMode for MC_BR_CrossCutterControl*)
	mcCUBIC_SPLINE : UINT := 256; (*interpolation rule*)
	mcCURRENT_DIR : USINT := 2; (*movement direction*)
	mcCYCLIC : UINT := 2; (*event move mode*)
	mcCYCLIC_ALL_EVENTS : UINT := 3; (*event move mode*)
	mcDATOBJ : UINT := 0; (*data object type*)
	mcDEFAULT_MOVE_PARAMETERS : INT := 1012; (*PLCopen motion parameter*)
	mcDIRECT : USINT := 7; (*start mode*)
	mcDIR_DEPENDENT : UINT := 1; (*mode for MPDC*)
	mcDIR_DEPENDENT_BACKLASH : UINT := 2; (*mode for MPDC*)
	mcDIR_DEPENDENT_SET_POSITION : UINT := 5; (*mode for MPDC*)
	mcDIR_INDEPENDENT : UINT := 3; (*mode for MPDC*)
	mcDIR_INDEPENDENT_SPEED : UINT := 4; (*mode for MPDC*)
	mcDISTANCE_BASED : UINT := 0; (*basis for cam movement (e.g. for MC_BR_CamTransition)*)
	mcDITHER : USINT := 32; (*setup mode*)
	mcEDGE_SENSITIVE : USINT := 4; (*additional mode for trigger event*)
	mcENABLE : UINT := 2;
	mcENABLE_LIMIT_NEG : INT := 5; (*PLCopen motion parameter*)
	mcENABLE_LIMIT_POS : INT := 4; (*PLCopen motion parameter*)
	mcENABLE_POS_LAG_MONITORING : INT := 6; (*PLCopen motion parameter*)
	mcENCODER : USINT := 0; (*setup mode*)
	mcENCODER_POSITION : UINT := 2; (*position source for MPDC*)
	mcEQUAL : UINT := 2;
	mcEVERY_RECORD : UINT := 1; (*mode for MC_BR_CyclicRead*)
	mcEXCEED_PERIOD : USINT := 8; (*movement direction*)
	mcFB_ERROR : USINT := 2;
	mcFB_INPUTS : REAL := 255.0; (*option for DefaultMoveParameters*)
	mcFF : USINT := 32; (*setup, torque mode*)
	mcFF_NEG_MOVE : UINT := 34; (*setup mode*)
	mcFF_POS_MOVE : UINT := 33; (*setup mode*)
	mcFILE : UINT := 1; (*data object type*)
	mcFILE_BIN : UINT := 0; (*binary format*)
	mcFILE_CSV : UINT := 1; (*CSV format*)
	mcFILE_TXT : UINT := 2; (*text format*)
	mcFIRST_RM : UINT := 0;
	mcFIRST_TRIGGER : UINT := 2;
	mcFLUX : USINT := 1; (*setup mode*)
	mcGE : UINT := 6;
	mcGET_BRAKE_STATUS : USINT := 16; (*brake command*)
	mcGREATER : UINT := 4;
	mcHARMONIC_COMBINATION : UINT := 8; (*motion rule*)
	mcHOLDOFF_DISTANCE : UINT := 16384;
	mcHOME_ABS_SWITCH : USINT := 2; (*homing mode*)
	mcHOME_ABSOLUTE : USINT := 4; (*homing mode*)
	mcHOME_ABSOLUTE_CORR : USINT := 6; (*homing mode*)
	mcHOME_AXIS_REF : USINT := 12; (*homing mode *)
	mcHOME_BLOCK_DS : USINT := 14; (*homing mode *)
	mcHOME_BLOCK_TORQUE : USINT := 13; (*homing mode *)
	mcHOME_DCM : USINT := 9; (*homing mode*)
	mcHOME_DCM_CORR : USINT := 10; (*homing mode*)
	mcHOME_DEFAULT : USINT := 0; (*homing mode*)
	mcHOME_DIRECT : USINT := 1; (*homing mode*)
	mcHOME_LIMIT_SWITCH : USINT := 3; (*homing mode*)
	mcHOME_REF_PULSE : USINT := 5; (*homing mode*)
	mcHOME_RESTORE_POS : USINT := 11; (*homing mode*)
	mcHOME_SET_PHASE : USINT := 7; (*homing mode*)
	mcHOME_SWITCH_GATE : USINT := 8; (*homing mode*)
	mcHORIZONTAL : USINT := 0; (*setup option for controller setup*)
	mcIDENTIFICATION : UINT := 10; (*setup mode *)
	mcIMMEDIATE : UINT := 0; (*mode for MC_BR_RegMarkCalc001, StartMode for MC_BR_CrossCutterControl, *)
	mcIN_WINDOW : USINT := 20; (*trigger event mode*)
	mcINC : USINT := 2; (*encoder type*)
	mcINC_ABS : USINT := 4; (*encoder type*)
	mcINC_REF : USINT := 3; (*encoder type*)
	mcINCLINED_SINE_CURVE : UINT := 5; (*motion rule*)
	mcINTERVAL_EVENT : UINT := 16;
    mcINVERSE : USINT := 255; (*encoder count direction*)
	mcIPL_LINEAR : USINT := 1; (*interpolation mode*)
	mcIPL_OFF : USINT := 0; (*interpolation mode*)
	mcIPL_QUADRATIC : USINT := 2; (*interpolation mode*)
	mcIPL_QUADRATIC_NO_OVERSHOOT : USINT := 4; (*interpolation mode*)
	mcISQ_F1_NOTCH : UINT := 128; (*setup mode*)
	mcISQ_F2_NOTCH : UINT := 256; (*setup mode*)
	mcISQ_F3_NOTCH : UINT := 512; (*setup mode*)
	mcISQ_RIPPLE : UINT := 20; (*setup mode*)
	mcLAST_POINT : UINT := 0; (*motion rule*)
	mcLEAD_IN : UINT := 2;
	mcLEAD_OUT : UINT := 4;
	mcLENGTH_ONLY : UINT := 32;
	mcLIMIT : USINT := 40; (*torque mode*)
	mcLIMIT_PARAMETERS : REAL := 1.0; (*option for DefaultMoveParameters*)
	mcLINEAR_CAM : USINT := 253; (*predefined 1:1 cam profile for MC_BR_CamDwell*)
	mcLINEAR_CAM_NON_PERIODIC : USINT := 254; (*for predifined 1:1 cam profile*)
	mcLINEAR_CAM_PERIODIC : USINT := 255; (*for predefined 1:1 cam profile*)
	mcLOAD : UINT := 276; (*trace command*)
	mcMANUAL_SEARCH : UINT := 64;
	mcMASTER_DISTANCE_BASED : UINT := 3; (*basis for movement profile (e.g. for MC_BR_Offset or MC_BR_Phasing)*)
    mcMASTER_INTERVAL : USINT := 0; (*start mode*)
	mcMASTER_POSITION : UINT := 256; (*additional basis for movement profile (e.g. for MC_BR_Offset), StartMode for MC_BR_CrossCutterControl*)
	mcMASTER_POSITION_BASED : UINT := 2; (*basis for movement profile (e.g. for MC_BR_Offset or MC_BR_Phasing)*)
	mcMAX_ACCELERATION_APPL : INT := 13; (*PLCopen motion parameter*)
	mcMAX_ACCELERATION_SYSTEM : INT := 12; (*PLCopen motion parameter*)
	mcMAX_DECELERATION_APPL : INT := 15; (*PLCopen motion parameter*)
	mcMAX_DECELERATION_SYSTEM : INT := 14; (*PLCopen motion parameter*)
	mcMAX_IV_TIME : USINT := 8; (*additional mode for power evaluation*)
	mcMAX_JERK : INT := 16; (*PLCopen motion parameter*)
	mcMAX_LOAD_SYSTEM : INT := 1015; (*PLCopen motion parameter*)
	mcMAX_POSITION_CHANGE : INT := 1016; (*PLCopen motion parameter*)
	mcMAX_POSITION_LAG : INT := 7; (*PLCopen motion parameter*)
	mcMAX_SLAVE_COMP_DISTANCE_NEG : UINT := 4; (*mode for automat compensation check*)
	mcMAX_SLAVE_COMP_DISTANCE_POS : UINT := 3; (*mode for automat compensation check*)
	mcMAX_VELOCITY_APPL : INT := 9; (*PLCopen motion parameter*)
	mcMAX_VELOCITY_SYSTEM : INT := 8; (*PLCopen motion parameter*)
	mcMIDDLE : USINT := 5;
	mcMIN_MASTER_COMP_DISTANCE : UINT := 2; (*mode for automat compensation check*)
	mcMODIFIED_ACCEL_TRAPEZOID : UINT := 6; (*motion rule*)
	mcMODIFIED_SINE_CURVE : UINT := 7; (*motion rule*)
	mcMOTOR : UINT := 258; (*switch on simulation mode*)
	mcMOVE_ACCELERATION_NEG : INT := 1005; (*PLCopen motion parameter*)
	mcMOVE_ACCELERATION_POS : INT := 1003; (*PLCopen motion parameter*)
	mcMOVE_CYCL_POS_IPL_MODE : INT := 1010; (*PLCopen motion parameter*)
	mcMOVE_CYCL_VEL_IPL_MODE : INT := 1011; (*PLCopen motion parameter*)
	mcMOVE_DECELERATION_NEG : INT := 1006; (*PLCopen motion parameter*)
	mcMOVE_DECELERATION_POS : INT := 1004; (*PLCopen motion parameter*)
	mcMOVE_VELOCITY_NEG : INT := 1002; (*PLCopen motion parameter*)
	mcMOVE_VELOCITY_POS : INT := 1001; (*PLCopen motion parameter*)
	mcMULTI_AXIS_TRACE : UDINT := 0; (*parameter trace type*)
	mcN_EDGE : USINT := 1;
	mcNEGATIVE_DIR : USINT := 1; (*movement direction*)
	mcNET_TRACE_GLOBAL : UDINT := 0; (*network trace type*)
	mcNETWORK_CYCLE_TIME: INT := 1017; (*PLCopen motion parameter*)
	mcNO_CHANGE_COMP : USINT := 2;
	mcNO_EVENTS : USINT := 253; (*event index*)
	mcNO_STATES : USINT := 253;
	mcNO_PARAMS : USINT := 253; (*parameter index*)
	mcNO_POSITION : USINT := 0;
	mcNO_START_COMP : USINT := 1;
	mcNO_TEXT : UINT := 0; (*no error text determination active*)
	mcNON_PERIODIC : BOOL := FALSE; (*cam profile mode*)
	mcNOT_AXIS_RELATED : UDINT := 16#FFFFFFFF;
	mcNULL : UINT := 1;
	mcOFF : BOOL := FALSE;
	mcON : BOOL := TRUE;
	mcONCE : UINT := 1;
	mcONE_RECORD : UINT := 0; (*mode for MC_BR_CyclicRead*)
	mcONLY_EVENTS : USINT := 254; (*event index*)
	mcONLY_PSM : USINT := 1; (*power evaluation  mode*)
	mcOPEN : USINT := 1;
	mcOPTIMIZED_ACCELERATION : UINT := 768; (*interpolation rule*)
	mcOPTIMIZED_VELOCITY : UINT := 512; (*interpolation rule*)
	mcOUT_WINDOW : USINT := 30; (*trigger event mode*)
	mcOVERRIDE : INT := 1000; (*PLCopen motion parameter*)
	mcP_EDGE : USINT := 0;
	mcPERIODIC : BOOL := TRUE; (*cam profile mode*)
	mcPOSITION : USINT := 1; (*setup mode*)
	mcPOSITIVE_DIR : USINT := 0; (*movement direction*)
	mcQUADRATIC_PARABOLA : UINT := 2; (*motion rule*)
	mcQUEUED : UINT := 1;
	mcRELATIVE : USINT := 1; (*start mode*)
	mcRELATIVE_NO_RESET : USINT := 3; (*start mode*)
	mcRESET : UINT := 320; (*trace command*)
	mcRESET_RING_STARTIDX : UINT := 4416; (*trace command (0x1000 + 0x0140)*)
	mcRESTART : UINT := 273; (*StartMode for MC_BR_CrossCutterControl*)
	mcREVERSE : UINT := 8;
	mcSATURATION : USINT := 30; (*setup mode*)
	mcSAVE : UINT := 341; (*trace command*)
	mcSAVE_RING_STARTIDX : UINT := 4437; (*trace command (0x1000 + 0x0155)*)
	mcSE : UINT := 3;
	mcSET_OFFSET : USINT := 34; (*setup mode*)
	mcSET_POSITION : UINT := 0; (*position source for MPDC*)
	mcSHIFT_FROM_EXPECTED : UINT := 50; (*input for MC_BR_TouchProbe*)
	mcSHIFT_FROM_RESULT : UINT := 49; (*input for MC_BR_TouchProbe*)
	mcSHORTEST_WAY : USINT := 3; (*synchronization mode, movement direction*)
	mcSIGNAL_CHIRP : UINT := 1; (*excitation signal type for controller setup*)
	mcSIGNAL_CHIRP_TRAPEZOID : UINT := 2; (*excitation signal type for controller setup*)
	mcSIGNAL_PRBS : UINT := 0; (*excitation signal type for controller setup*)
	mcSIMPLE_SINE_CURVE : UINT := 3; (*motion rule*)
	mcSIMULATION_INIT : UINT := 512; (*initialize simulation parameters*)
	mcSIMULATION_OFF : UINT := 259; (*switch off simulation mode*)
	mcSIMULATION_ON : UINT := 258; (*switch on simulation mode*)
	mcSIMULATION_READ : UINT := 265; (*read calculated simulation parameters*)
	mcSLAVE_POSITION : UINT := 0; (*additional basis for movement profile (e.g. for MC_BR_Offset)*)
	mcSLOW_DOWN : USINT := 5; (*synchronization mode*)
	mcSMALLER : UINT := 1;
	mcSPEED : USINT := 2; (*setup mode*)
    mcSTANDARD : USINT := 0; (*encoder count direction*)
	mcSTART : UINT := 260;
	mcSTART_N_FLANK : UINT := 128; (*start MPDC at negative flank*)
	mcSTART_ONLY : USINT := 3; (*power evaluation mode*)
	mcSTART_P_FLANK : UINT := 0; (*start MPDC at positive flank*)
	mcSTEPPER : USINT := 31; (*setup mode*)
	mcSTOP : UINT := 261;
	mcSTOP_INDEX : INT := 1013; (*PLCopen motion parameter*)
	mcSTRAIGHT_LINE : UINT := 1; (*motion rule*)
	mcSW_END_ACTIVE : REAL := 0.0; (*SW end monitoring mode*)
	mcSW_END_IGNORE : REAL := 1.0; (*SW end monitoring mode*)
	mcSW_END_MONITORING : INT := 1014; (*PLCopen motion parameter*)
	mcSW_END_SPF : REAL := 2.0; (*SW end monitoring mode*)
	mcSW_LIMIT_NEG : INT := 3; (*PLCopen motion parameter*)
	mcSW_LIMIT_POS : INT := 2; (*PLCopen motion parameter*)
	mcSWITCH_OFF : UINT := 259; (*trace command*)
	mcSWITCH_ON : UINT := 258; (*trace command*)
	mcT_FILTER : UINT := 64; (*setup mode*)
	mcT_FILTER_2 : UINT := 65; (*setup mode*)
	mcTEST : UINT := 31; (*setup mode*)
	mcTEXT : UINT := 1; (*error text determination active*)
	mcTIME_BASED : UINT := 1; (*basis for movement profile (e.g. for MC_BR_Offset or MC_BR_Phasing)*)
	mcTIME_LIMIT : USINT := 8; (*enable time dependent switch off of function*)
	mcTRACE_DELAY : USINT := 6; (*trace status*)
	mcTRACE_FINISHED : USINT := 1; (*trace status*)
	mcTRACE_REST : USINT := 5; (*trace status*)
	mcTRACE_RING : USINT := 4; (*trace status*)
	mcTRACE_STARTED : USINT := 20; (*trace status*)
	mcTRACE_TIME : USINT := 2; (*trace status*)
	mcTRACE_TRIGGER : USINT := 3; (*trace status*)
	mcTRANSITION_OFF : UINT := 0;
	mcTRANSITION_ON : UINT := 1;
	mcTUNE_STANDSTILL : USINT := 0; (*constant for OperatingPoint*)
    mcTUNE_TN : UINT := 16; (*setup mode*)
	mcTUNE_V_CONSTANT : USINT := 1; (*constant for OperatingPoint*)
	mcUNEQUAL : UINT := 5;
	mcUPDATE_PERIOD : UINT := 16#8000; (*input for MC_BR_TouchProbe*)
	mcUSE_AXIS_PERIOD : UINT := 16#4000; (*input for MC_BR_TouchProbe*)
	mcUSE_FILTER_PAR : UINT := 4; (*setup mode *)
	mcUSE_FIRST_TRIGGER_POS : UINT := 64; (*additional input for MC_BR_TouchProbe*)
	mcUSE_STOP_COMP : USINT := 4;
	mcUSE_TN : UINT := 8; (*setup mode*)
	mcV_LIMIT_CALC : USINT := 4; (*recalculate speed limit depending on user setting*)
	mcV_LIMIT_OFF : USINT := 2; (*disable speed limit*)
	mcVELOCITY_CONTROL : UINT := 4; (*basis for movement profile (e.g. for MC_BR_Offset or MC_BR_Phasing)*)
	mcVERTICAL : USINT := 1; (*setup option for controller setup*)
	mcWITH_PARAM : USINT := 2; (*power evaluation mode*)
	mcWITHIN_PERIOD : USINT := 6; (*synchronization mode*)
	mcWITHOUT_PERIOD : UINT := 4; (*input for MC_BR_TouchProbe*)
	mcWITH_FF : USINT := 0; (*torque limit mode*)
	mcWITHOUT_FF : USINT := 1; (*torque limit mode*)
	mcWRAP : UINT := 2;
	mcWRITE_DIRECT : UINT := 256; (*cyclic write mode*)
END_VAR
